(* IEC 61131-3 sources: daoli-st-library/DL_Device (part 17) *)

(* ---- FB_DL_CombinerArcDetect.st ---- *)
(*
  FB_DL_CombinerArcDetect  —  汇流箱直流拉弧特征判据 / Combiner box DC arc feature detection
  分类 Category : DL_Device
  码位 Code     : 16#03_2_00
  版本 Version  : 1.0.1
  溯源 Source   : NAMUR NE107 语义借鉴 · clean-room 实现，仅借分类/参数域/命名，未复制源码
  修订 Revision : v1.0.1 (R34 终审抽检) — ① 段 1 复位只清组态码 16#0002_0300，不再连带清 16#0002_0310
                  （原「无条件清锁存」使拉弧仍在时 bError 掉为 FALSE、uErrorId 归 0，而 eNe107 仍报 eFailure，
                  故障位/事件码/NE107 三者不同步，且 eAlarm 解除需第二次复位沿）；
                  ② bCfgOk 补 tSampleTime / tFilterTC 正域闸（原 0 或负值时高通静默不动作、永不告警，违 R179）。
                  接口、码表、NE107 映射不变。
  功能 Function : 1) 高通滤波提取电流高频分量，超门限按多拍持续确认才升故障（单拍尖峰只计信息级）；
                  2) 采样率与滤波截止频率配比校验（截止 >= 采样率/2 即出厂报码，不进入判据）；
                  3) 分级出口按 NE107 六态映射，未知态归 eUnknown 绝不归 eOk。
  边界 Boundary : ① 高频分量提取前确认采样率/截止频率配比合法（截止 >= 采样率/2 即报码）；
                  ② 拉弧判据多拍持续确认，单拍尖峰只计信息级不升故障；
                  ③ 分级出口按 NE107 六态映射，未知态归 eUnknown（不归 eOk）；
                  ④ 输出三行同向：高频分量 → 确认计数 → 拉弧标志。
  依赖 Depends  : FB_DL_HighPassFilter（高频分量提取，每拍无条件调用）

  码表 Error codes（本件子码步进 16#10，避让邻件码位）:
    16#0002_0300 故障级：采样率/截止频率配比非法（截止 >= 采样率/2）或采样率 <= 0
    16#0002_0310 故障级：拉弧已确认（多拍持续超门限），需 bReset 清除
    16#0002_0320 信息级：单拍尖峰（未达确认拍数，不置 bError）
*)

TYPE E_DL_CadNe107 :
(
    eOk                  := 0,   // 正常 / Normal
    eFailure             := 10,  // 故障 / Failure
    eCheckFunction       := 20,  // 功能检查 / Function check
    eOutOfSpec           := 30,  // 超出规格 / Out of specification
    eMaintenanceRequired := 40,  // 需要维护 / Maintenance required
    eUnknown             := 90   // 未知态（兜底）/ Unknown fallback
);
END_TYPE

TYPE E_DL_CadPhase :
(
    eIdle    := 0,   // 空闲 / Idle
    eWatch   := 10,  // 常规监视 / Normal watch
    eConfirm := 20,  // 多拍确认中 / Multi-scan confirmation
    eAlarm   := 30,  // 拉弧告警 / Arc alarm
    eFault   := 90   // 组态故障锁定 / Configuration fault locked
);
END_TYPE

FUNCTION_BLOCK FB_DL_CombinerArcDetect
VAR_INPUT
    bEnable       : BOOL;                         // 总使能，FALSE 回空闲 / Master enable
    bReset        : BOOL;                          // 复位，上升沿清告警与故障 / Reset
    fCurrentA     : REAL;                         // 直流支路电流 [A]，域 0~30 / DC branch current [A]
    fSampleRateHz : REAL := 10000.0;              // 电流采样率 [Hz]，域 > 0 / Current sampling rate [Hz]
    fCutoffHz     : REAL := 2000.0;               // 高通截止频率 [Hz]，须 < 采样率/2 / High-pass cutoff [Hz]
    fHfThreshA    : REAL := 0.15;                 // 高频分量门限 [A]，域 > 0 / HF component threshold [A]
    nConfirmScans : INT := 5;                     // 持续确认拍数 [拍]，域 1~100 / Confirmation scans, 1..100
    tFilterTC      : TIME := T#20MS;              // 高通时间常数 [ms] / High-pass time constant [ms]
    tSampleTime   : TIME := T#10MS;               // 任务采样周期 [ms]，域 > 0 / Task sample period [ms]
    fEps          : REAL := 1.0E-6;               // 浮点判零容差 [1] / Floating zero tolerance
END_VAR
VAR_OUTPUT
    fHfOutA       : REAL;                         // 高频分量输出 [A] / HF component output [A]
    nConfirmCnt   : INT;                          // 当前确认计数 [拍] / Current confirmation counter
    bArcAlarm     : BOOL;                         // 拉弧告警（保持型）/ Arc alarm, held
    bSpikeOnly    : BOOL;                         // 仅单拍尖峰（信息级）/ Single-scan spike only
    eNe107        : E_DL_CadNe107;                // NE107 六态映射出口，段尾单点赋值 / NE107 mapping, single write
    bError        : BOOL;                         // 故障标志，与故障级码配对 / Fault flag paired with fault codes
    uErrorId      : UDINT;                        // 事件码，0 = 无事件 / Event code, 0 = none
    eStateOut     : E_DL_CadPhase;                // 状态机当前态，段尾单点映射 / Phase mapped at tail
END_VAR
VAR
    _eState       : E_DL_CadPhase := E_DL_CadPhase.eIdle;  // 内部状态 / Internal state
    rtrReset      : R_TRIG;                       // 复位沿 / Reset edge
    fbHp          : FB_DL_HighPassFilter;         // 高通滤波实例（无条件调用）/ High-pass filter instance
    bCfgOk        : BOOL;                         // 配比组态合法 / Ratio configuration valid
    bSigOk        : BOOL;                         // 电流采样有效 / Current sample valid
    bOver         : BOOL;                         // 本拍超门限 / Over threshold this scan
    nCnt          : INT;                          // 确认计数暂存 [拍] / Confirmation counter buffer
    eMap          : E_DL_CadNe107;                // NE107 映射暂存（单点写入源）/ NE107 mapping buffer
    uFault        : UDINT;                        // 锁存故障码 / Latched fault code
    uInfo         : UDINT;                        // 信息级码 / Information code
END_VAR
VAR CONSTANT
    DL_CAD_CNTMAX : INT := 1000;                  // 确认计数上限 [拍]，防溢出 / Confirmation counter ceiling
    DL_CAD_SRMAX  : REAL := 1.0E6;                // 采样率物理域上限 [Hz] / Sampling rate domain high
END_VAR

(* === 段 0 · 实例刷新（无条件周期调用）=== *)
rtrReset(CLK := bReset);                          // 每拍刷新复位沿

(* === 段 1 · 组态闸：采样率/截止频率配比（截止 >= 采样率/2 即报码）=== *)
bCfgOk := (fSampleRateHz > fEps) AND (fSampleRateHz <= DL_CAD_SRMAX)
          AND (fCutoffHz > fEps)
          AND (fCutoffHz < (fSampleRateHz * 0.5))          // Nyquist 配比硬判据
          AND (fHfThreshA > fEps) AND (nConfirmScans >= 1) AND (nConfirmScans <= 100)
          AND (TIME_TO_LREAL(tSampleTime) > 0.0) AND (TIME_TO_LREAL(tFilterTC) > 0.0)   // 节拍/时间常数正域闸（R179）
          AND (fSampleRateHz = fSampleRateHz) AND (fCutoffHz = fCutoffHz)
          AND (fHfThreshA = fHfThreshA);                   // 含 NaN 自反判据
IF NOT bCfgOk THEN
    uFault := 16#0002_0300;                       // 故障级：配比非法
END_IF
IF rtrReset.Q AND bCfgOk THEN
    IF uFault <> 16#0002_0310 THEN
        uFault := 16#0000;                        // 复位沿清锁存（拉弧码由 eAlarm 相专清，保持位码同步）
    END_IF
    IF NOT bArcAlarm THEN
        nCnt := 0;                                // 未进入告警时清确认计数
    END_IF
END_IF
bSigOk := (fCurrentA = fCurrentA) AND (ABS(fCurrentA) < 1.0E30) AND (fCurrentA >= 0.0);   // NaN 自反 + 域闸
uInfo := 16#0000;                                 // 信息码每拍清零

(* === 段 2 · 高频分量实例（每拍无条件调用）=== *)
fbHp(bEnable := bEnable AND bSigOk AND bCfgOk,    // 配比非法/信号无效时不使能（禁误判）
     fIn := fCurrentA,                            // 电流采样
     tTimeConst := tFilterTC,                     // 高通时间常数
     tSampleTime := tSampleTime,                  // 采样周期
     rOutMin := -1000.0,                          // 输出下限 [A]
     rOutMax := 1000.0,                           // 输出上限 [A]
     bTrack := rtrReset.Q,                        // 复位沿清基线
     fTrackValue := 0.0);                         // 跟踪值 0
fHfOutA := fbHp.fOut;                             // 高频分量输出
bOver := bCfgOk AND bSigOk AND fbHp.bValid AND (ABS(fHfOutA) >= fHfThreshA);   // 超门限判据

(* === 段 3 · 主状态机（ENUM + CASE，含 ELSE 兜底）=== *)
CASE _eState OF
E_DL_CadPhase.eIdle :
    nCnt := 0;                                    // 空闲计数清零
    bSpikeOnly := FALSE;                          // 尖峰标志复位
    IF uFault = 16#0002_0300 THEN
        _eState := E_DL_CadPhase.eFault;          // 组态故障优先
    ELSIF bEnable AND bCfgOk THEN
        _eState := E_DL_CadPhase.eWatch;          // 进入监视相
    END_IF

E_DL_CadPhase.eWatch :
    IF bOver THEN
        nCnt := 1;                                // 首拍超门限：进入确认
        _eState := E_DL_CadPhase.eConfirm;
    ELSE
        IF bSpikeOnly THEN
            uInfo := 16#0002_0320;                // 信息级：单拍尖峰记录（不升故障）
        END_IF
        bSpikeOnly := bSpikeOnly AND bOver;       // 无超门限拍则尖峰记录清除
    END_IF

E_DL_CadPhase.eConfirm :
    IF bOver THEN
        nCnt := nCnt + 1;                         // 连续超门限：计数累加
        IF nCnt > DL_CAD_CNTMAX THEN
            nCnt := DL_CAD_CNTMAX;                // 饱和防溢出
        END_IF
        IF nCnt >= nConfirmScans THEN
            bArcAlarm := TRUE;                    // 置位型：拉弧确认告警（段尾不清零）
            uFault := 16#0002_0310;               // 故障级：拉弧已确认
            _eState := E_DL_CadPhase.eAlarm;      // 转告警相
        END_IF
    ELSE
        bSpikeOnly := TRUE;                       // 未达确认拍数即回落：只计单拍尖峰
        uInfo := 16#0002_0320;                    // 信息级：单拍尖峰
        nCnt := 0;                                // 计数清零（要求连续）
        _eState := E_DL_CadPhase.eWatch;          // 回监视相
    END_IF

E_DL_CadPhase.eAlarm :
    bArcAlarm := TRUE;                            // 告警保持
    IF NOT bOver AND rtrReset.Q THEN
        uFault := 16#0000;                        // 超门限消失且复位沿：清锁存
        bArcAlarm := FALSE;                       // 告警解除（可到达的解除路径）
        nCnt := 0;                                // 计数清零
        _eState := E_DL_CadPhase.eWatch;
    END_IF

E_DL_CadPhase.eFault :
    nCnt := 0;                                    // 故障态计数清零
    bArcAlarm := FALSE;                           // 故障态不告警（配置错误优先）
    IF uFault = 16#0000 THEN
        _eState := E_DL_CadPhase.eIdle;           // 解锁回空闲
    END_IF

ELSE
    _eState := E_DL_CadPhase.eFault;              // 非法状态拦截
    uFault := 16#0002_0300;                       // 故障级：相 ID 越界
    bArcAlarm := FALSE;                           // 安全侧不告警
END_CASE
IF NOT bEnable THEN
    _eState := E_DL_CadPhase.eIdle;               // 失能最高优先回空闲
    bArcAlarm := FALSE;                           // 失能清告警
    nCnt := 0;                                    // 失能清计数
    IF uFault = 16#0002_0310 THEN
        uFault := 16#0000;                        // 失能同拍清拉弧锁存：相序丢失后 eAlarm 不可达，防锁死（终审式 1）
    END_IF
END_IF

(* === 段 4 · 输出映射与 NE107 六态（段尾单点赋值）=== *)
nConfirmCnt := nCnt;                              // 确认计数输出
CASE _eState OF
E_DL_CadPhase.eWatch :
    eMap := E_DL_CadNe107.eOk;                    // 常规监视：正常态
E_DL_CadPhase.eConfirm :
    eMap := E_DL_CadNe107.eMaintenanceRequired;   // 确认中：需维护关注
E_DL_CadPhase.eAlarm :
    eMap := E_DL_CadNe107.eFailure;               // 拉弧确认：故障态
E_DL_CadPhase.eFault :
    eMap := E_DL_CadNe107.eOutOfSpec;             // 组态越规格
E_DL_CadPhase.eIdle :
    eMap := E_DL_CadNe107.eCheckFunction;         // 空闲未监视：功能检查
ELSE
    eMap := E_DL_CadNe107.eUnknown;               // 未知态兜底：绝不归 eOk
END_CASE
IF bSpikeOnly AND (eMap = E_DL_CadNe107.eOk) THEN
    eMap := E_DL_CadNe107.eMaintenanceRequired;   // 单拍尖峰：提升到需维护（信息级）
END_IF
eNe107 := eMap;                                   // 单点写入 NE107 出口
bError := (uFault <> 16#0000);                    // 故障标志仅由故障级码置位（R45 配对）
IF bError THEN
    uErrorId := uFault;                           // 故障级优先上报
ELSE
    uErrorId := uInfo;                            // 否则上报信息级码
END_IF
eStateOut := _eState;                             // 输出枚举段尾单点映射（N2 规则）
END_FUNCTION_BLOCK

(* ---- FB_DL_CondensateDrainSeq.st ---- *)
(*
  ==================================================================
  组件名 Component  : FB_DL_CondensateDrainSeq
  分类   Category   : DL_Device
  复杂度 Complexity  : cx5
  版本   Version    : 1.0.0
  功能   Purpose    : 储气罐 / 空压机冷凝水自动排污阀时序。定时触发与液位高
                      双触发源并联起排；开阀确认反馈 → 排放（触发消失且最
                      小排放时长满足）→ 关阀确认反馈；三窗超时诊断（开阀 /
                      排放 / 关阀独立成因独立码位语义，R190）。
  来源   Source     : t2-2-lbp（命令→监视→判定三段）
  溯源   Origin     : IEC 61131-3 标准语义的道莅防御性实现；冷凝水排污双触
                      发与阀反馈确认窗为行业公知工程语义，clean-room 自研实
                      现，未复制 LBP 或任何厂商私有库源码。
  平台   Platform   : 纯 IEC 61131-3（Standard.library: TON / R_TRIG，无私有库）
  分工声明 Split     : 与 DL_Device 存量阀类执行件（电磁阀直控类）分工——直
                      控件只做单阀开关映射，本件为排污全过程顺控（三窗监视
                      与诊断）；不做压力 / 温度工艺调节。
  作者   Author     : 道莅代码库 · PLC 编程专家（R58）
  ------------------------------------------------------------------
  边界 Boundary     :
                      一 组态配比约束（R100）：tMinDrain < tDrainMax（最小排
                         放短于排放超时）且 tOpenConfirm > T#0S 且 tCloseConfirm
                         > T#0S；越域判故障级锁存；
                      二 触发为电平语义：定时触发与液位高任一为真且许可满
                         足即起排；排放相退出 = 触发消失（事件）AND 最小排放
                         时长满足（双条件，R98 精神）；
                      三 故障相阀命令安全侧断开（排污阀断电 = 关闭，R191 显
                         式声明）；故障锁存解除路径 = bReset 上升沿（唯一路
                         径，R188）；
                      四 无全局变量、无外部变量声明、无物理地址寻址。
  修订记录 Revision  :
    2026-11-21  v1.0.0  R58 首版（批 3 · 序号 11）
  ==================================================================
*)

TYPE E_DL_CdsPhase :
(
    eCdsIdle    := 0,  // 空闲：等触发 / idle, waiting for a trigger
    eCdsOpening := 10, // 开阀：等阀开反馈确认 / opening, awaiting the open feedback
    eCdsDraining := 20, // 排放中：等触发消失且最小时长满足 / draining, awaiting the trigger gone with the minimum met
    eCdsClosing := 30, // 关阀：等阀关反馈确认 / closing, awaiting the closed feedback
    eCdsFault   := 90  // 故障锁存 / the latched fault
);
END_TYPE

TYPE E_DL_CdsCause :
(
    eNone         := 0, // 无成因 / no cause
    eCfgBad       := 1, // 组态非法：时间窗配比越域（故障级，与 bError 配对）/ an illegal config
    eValveOpenTo  := 2, // 开阀确认超时（故障级，与 bError 配对）/ an open confirm timeout
    eDrainTimeout := 3, // 排放超时（液位不回落，故障级，与 bError 配对）/ a drain timeout
    eValveCloseTo := 4, // 关阀确认超时（故障级，与 bError 配对）/ a close confirm timeout
    ePhaseBad     := 5  // 非法相位兜底（故障级，与 bError 配对）/ an illegal phase fallback
);
END_TYPE

FUNCTION_BLOCK FB_DL_CondensateDrainSeq
VAR_INPUT
    bEnable       : BOOL := TRUE;   // 使能，失能回空闲关阀 [-] / enable, disabling returns idle with the valve closed
    bReset        : BOOL := FALSE;  // 复位上升沿清故障锁存 [-] / reset rising edge clears the latch
    bTimTrig      : BOOL := FALSE;  // 定时触发电平（调用方定时器给出）[-] / the timer trigger level
    bLevelHigh    : BOOL := FALSE;  // 液位高触发电平 [-] / the level high trigger level
    bPermitDrain  : BOOL := TRUE;   // 排放许可（压力低联锁给出）[-] / the drain permit from the pressure interlock
    bFbValveOpen  : BOOL := FALSE;  // 排污阀开到位反馈 [-] / the valve open feedback
    bFbValveClosed: BOOL := TRUE;   // 排污阀关到位反馈 [-] / the valve closed feedback
    tOpenConfirm  : TIME := T#5S;   // 开阀确认窗 [毫秒] / the open confirm window [millisecond]
    tDrainMax     : TIME := T#60S;  // 排放超时窗 [毫秒] / the drain timeout window [millisecond]
    tCloseConfirm : TIME := T#5S;   // 关阀确认窗 [毫秒] / the close confirm window [millisecond]
    tMinDrain     : TIME := T#2S;   // 最小排放时长 [毫秒] / the minimum drain duration [millisecond]
END_VAR
VAR_OUTPUT
    bValveCmd   : BOOL := FALSE; // 排污阀命令输出（TRUE = 开阀）[-] / the valve command outlet, true = open
    bDrainActive: BOOL := FALSE; // 排放进行指示 [-] / the drain active indicator
    ePhase      : E_DL_CdsPhase := E_DL_CdsPhase.eCdsIdle; // 相位出口 [枚举] / the phase outlet
    eCause      : E_DL_CdsCause := E_DL_CdsCause.eNone; // 成因出口，锁存回放 [枚举] / the cause outlet replayed
    bError      : BOOL := FALSE; // 故障锁存标志 [-] / the fault latch flag
END_VAR
VAR
    rtReset : R_TRIG; // 复位沿检测，段 0 无条件刷新 / the reset edge
    tonOpen : TON;    // 开阀确认窗，段 0 无条件刷新 / the open confirm window
    tonDrain: TON;    // 排放超时窗，段 0 无条件刷新 / the drain timeout window
    tonClose: TON;    // 关阀确认窗，段 0 无条件刷新 / the close confirm window
    tonMin  : TON;    // 最小排放窗，段 0 无条件刷新 / the minimum drain window
    _ePhase : E_DL_CdsPhase := E_DL_CdsPhase.eCdsIdle; // 内部相位，CASE 唯一写入目标 / the internal phase
    _eFaulC : E_DL_CdsCause := E_DL_CdsCause.eNone; // 故障级成因，锁存至复位沿 / the fault cause latched
    _bFault : BOOL := FALSE; // 故障锁存位 [-] / the fault latch bit
    _bCfgOk : BOOL := FALSE; // 组态域内 [-] / the config inside the domain
    _bInit  : BOOL := FALSE; // 首扫初始化完成标志（R310）/ the first scan flag
END_VAR

// 段 0｜定时器与沿检测无条件周期刷新（禁入分支，FB50-1）/ segment 0, the unconditional refresh
rtReset(CLK := bReset); // 复位沿 / the reset edge
tonOpen(IN := (_ePhase = E_DL_CdsPhase.eCdsOpening) AND (NOT _bFault) AND bEnable, PT := tOpenConfirm); // 开阀窗，IN 串开阀相闸 / the open window gated by the opening phase
tonDrain(IN := (_ePhase = E_DL_CdsPhase.eCdsDraining) AND (NOT _bFault) AND bEnable, PT := tDrainMax); // 排放窗，IN 串排放相闸 / the drain window gated by the draining phase
tonClose(IN := (_ePhase = E_DL_CdsPhase.eCdsClosing) AND (NOT _bFault) AND bEnable, PT := tCloseConfirm); // 关阀窗，IN 串关阀相闸 / the close window gated by the closing phase
tonMin(IN := (_ePhase = E_DL_CdsPhase.eCdsDraining) AND (NOT _bFault) AND bEnable, PT := tMinDrain); // 最小排放窗，与排放窗同相起算（配比约束见边界一）/ the minimum window co-started with the drain window

// 段 1｜首扫初始化（R310）/ segment 1, the first scan
IF NOT _bInit THEN // 首扫一拍 / the first scan
    _bInit := TRUE; // 置首扫标志 / raise the flag
END_IF

// 段 2｜复位沿作用域：清故障锁存 / 迁空闲（两项逐项声明，边界三）/ segment 2, the reset edge scope
IF rtReset.Q THEN // 复位沿 / the reset edge
    _bFault := FALSE; // 作用域一：清故障锁存 / scope one, clear the fault latch
    _eFaulC := E_DL_CdsCause.eNone; // 作用域一：清成因 / scope one, clear the cause
    _ePhase := E_DL_CdsPhase.eCdsIdle; // 作用域二：迁空闲相 / scope two, back to idle
END_IF

// 段 3｜组态域闸（边界一，R100 配比）/ segment 3, the config gate
_bCfgOk := (tOpenConfirm > T#0S) AND (tCloseConfirm > T#0S) AND (tMinDrain < tDrainMax) AND (tDrainMax > T#0S); // 确认窗 / 排放窗 / 配比判定 / the confirm, drain and pairing verdicts
IF NOT _bCfgOk THEN // 配比越域 / a pairing violation
    IF NOT _bFault THEN // 未锁存才迁移 / migrate only while unlatched
        _bFault := TRUE; // 置故障锁存 / raise the fault latch
        _eFaulC := E_DL_CdsCause.eCfgBad; // 故障级成因（R45 配对）/ the fault cause
        _ePhase := E_DL_CdsPhase.eCdsFault; // 迁故障相（锁存与迁相同分支，FB50-1）/ migrate to the fault phase
    END_IF
END_IF

// 段 4｜相位机：ENUM + CASE，含 ELSE 非法相位兜底（R128）/ segment 4, the phase machine
CASE _ePhase OF

E_DL_CdsPhase.eCdsIdle: // 空闲相：双触发源并联评估（边界二）/ the idle phase, the dual trigger evaluation
    IF NOT bEnable THEN // 失能驻留 / dwell while disabled
        _ePhase := E_DL_CdsPhase.eCdsIdle; // 停摆驻留 / dwell
    ELSIF (bTimTrig OR bLevelHigh) AND bPermitDrain THEN // 触发且许可 / a trigger with the permit
        _ePhase := E_DL_CdsPhase.eCdsOpening; // 迁开阀相 / migrate to the opening phase
    END_IF

E_DL_CdsPhase.eCdsOpening: // 开阀相：等阀开反馈确认 / the opening phase
    IF NOT bEnable THEN // 失能回空闲关阀（R191 显式）/ a disable returns idle
        _ePhase := E_DL_CdsPhase.eCdsIdle; // 回空闲相 / back to idle
    ELSIF bFbValveOpen THEN // 阀开反馈确认 / the open feedback confirmed
        _ePhase := E_DL_CdsPhase.eCdsDraining; // 迁排放相 / migrate to the draining phase
    ELSIF tonOpen.Q THEN // 开阀确认窗超时（R190 独立成因）/ the open timeout, an independent cause
        _bFault := TRUE; // 置故障锁存 / raise the fault latch
        _eFaulC := E_DL_CdsCause.eValveOpenTo; // 故障级成因（R45 配对）/ the fault cause
        _ePhase := E_DL_CdsPhase.eCdsFault; // 迁故障相 / migrate to the fault phase
    END_IF

E_DL_CdsPhase.eCdsDraining: // 排放相：双退出条件（边界二，R98 精神）/ the draining phase, the dual exit
    IF NOT bEnable THEN // 失能回空闲关阀 / a disable returns idle
        _ePhase := E_DL_CdsPhase.eCdsIdle; // 回空闲相 / back to idle
    ELSIF (NOT bTimTrig) AND (NOT bLevelHigh) AND tonMin.Q THEN // 触发消失且最小排放时长满足 / the trigger gone with the minimum met
        _ePhase := E_DL_CdsPhase.eCdsClosing; // 迁关阀相 / migrate to the closing phase
    ELSIF tonDrain.Q THEN // 排放超时（液位不回落，R190 独立成因）/ the drain timeout, an independent cause
        _bFault := TRUE; // 置故障锁存 / raise the fault latch
        _eFaulC := E_DL_CdsCause.eDrainTimeout; // 故障级成因（R45 配对）/ the fault cause
        _ePhase := E_DL_CdsPhase.eCdsFault; // 迁故障相 / migrate to the fault phase
    END_IF

E_DL_CdsPhase.eCdsClosing: // 关阀相：等阀关反馈确认 / the closing phase
    IF NOT bEnable THEN // 失能回空闲 / a disable returns idle
        _ePhase := E_DL_CdsPhase.eCdsIdle; // 回空闲相 / back to idle
    ELSIF bFbValveClosed THEN // 阀关反馈确认 / the closed feedback confirmed
        _ePhase := E_DL_CdsPhase.eCdsIdle; // 回空闲相 / back to idle
    ELSIF tonClose.Q THEN // 关阀确认窗超时（R190 独立成因）/ the close timeout, an independent cause
        _bFault := TRUE; // 置故障锁存 / raise the fault latch
        _eFaulC := E_DL_CdsCause.eValveCloseTo; // 故障级成因（R45 配对）/ the fault cause
        _ePhase := E_DL_CdsPhase.eCdsFault; // 迁故障相 / migrate to the fault phase
    END_IF

E_DL_CdsPhase.eCdsFault: // 故障相：成因锁存等复位沿；阀命令安全侧断开 / the fault phase
ELSE // 非法相位兜底（R128）/ the illegal phase fallback
    _bFault := TRUE; // 置故障锁存 / raise the fault latch
    _eFaulC := E_DL_CdsCause.ePhaseBad; // 故障级成因（R45 配对）/ the fault cause
    _ePhase := E_DL_CdsPhase.eCdsFault; // 迁故障相 / migrate to the fault phase
END_CASE

// 段 5｜统一出口（边界三安全侧）/ segment 5, the unified outlet
bValveCmd := ((_ePhase = E_DL_CdsPhase.eCdsOpening) OR (_ePhase = E_DL_CdsPhase.eCdsDraining)) AND bEnable AND (NOT _bFault); // 阀命令仅开阀与排放相 / the valve command in the opening and draining phases
bDrainActive := (_ePhase = E_DL_CdsPhase.eCdsDraining) AND (NOT _bFault); // 排放指示 / the drain indicator
ePhase := _ePhase; // 相位出口单点映射 / the phase outlet
IF _bFault THEN // 故障锁存优先 / the fault latch first
    eCause := _eFaulC; // 成因锁存回放（R152）/ the cause replayed
ELSE // 无锁存 / no latch
    eCause := E_DL_CdsCause.eNone; // 无成因 / no cause
END_IF
bError := _bFault; // 故障标志与锁存位同源 / the flag shares the latch
END_FUNCTION_BLOCK

(* ---- FB_DL_ContactorWeldDetect.st ---- *)
(*==============================================================================
 * 组件名称 (Component)  : FB_DL_ContactorWeldDetect
 * 所属子库 (Sublibrary) : DL_Device
 * 当前版本 (Version)    : 1.0.0
 * 兼容性   (Platform)   : CODESYS 3.5+ / TwinCAT 3 / 汇川 InoProShop / 施耐德 Machine Expert
 *                         仅依赖 Standard.library（TON / R_TRIG）与库内健康枚举唯一属主，
 *                         零厂商私有库
 * 功能描述 (Function)   : 接触器熔焊与不吸合检测。① 熔焊：断开指令后 tReleaseMax 内反馈仍为 1
 *                         → eCause = eWeld，故障锁存；② 不吸合：闭合指令后 tPickupMax 内无反馈
 *                         → eCause = eNoPickup，故障锁存。两成因各有独立 TON 与独立归因成员
 *                         （R190 归因唯一，禁止共用一个成因导致另一端永不赋值）。
 * 复位语义 (Design)     : **熔焊为不可自恢复故障**：解除式要求「复位沿 ∧ 反馈已回落」。若反馈是
 *                         真实熔焊，反馈不会回落 → 复位**不解锁**，这是**设计意图**而非缺陷：
 *                         触点焊死时允许软复位等于给现场一个「假修复」通道，会把带电粘连的
 *                         主回路重新投入。现场处置只能是更换接触器后反馈自然回落再复位。
 * 归属声明 (Ownership)  : 健康出口 eHealth 引用枚举 `E_DL_Ne107Status` 唯一属主，属主文件为
 *                         `C:\Library\DL_Device\I_DL_DeviceHealth.st`（枚举定义位于该文件 L91 附近），
 *                         本件只引用不重复声明（全库同名枚举定义计数 = 1，R67）。
 * 接口     (Interface)  : 输入 bCmdClose 闭合指令、bFbClosed 触点反馈、tReleaseMax 释放超时、
 *                         tPickupMax 吸合超时、bReset 复位；输出 bWeldSuspect 熔焊疑似位、
 *                         eCause 归因、eHealth NE107 健康态、eState / bError / nErrId。
 * 边界     (Boundary)   : ① 组态闸：tReleaseMax <= T#0S 或 tPickupMax <= T#0S → 故障锁存；
 *                         ② TON 两枚 + R_TRIG 一枚段 0 无条件周期刷新，IN 由当拍指令与反馈派生；
 *                         ③ 故障相迁出唯一路径 = bReset 上升沿；④ 零全局耦合（无 GVL / 无物理地址）。
 * 解除式   (Release)    : bReset 上升沿 ∧ 组态合法 ∧ 反馈已回落（bFbClosed = FALSE，当拍量，
 *                         R240 范式）。自证可满足（终审两式 1）：反馈为真实熔焊时该式不可满足，
 *                         属刻意的安全不可解除；触点更换后反馈回落即达，故路径物理可达。
 * 码表     (Codes)      : 16#0003_0702 故障级：接触器故障总码（组态非法 / 熔焊 / 不吸合 / 非法相位），
 *                         锁存至 bReset 上升沿，归因由 eCause 承载（R190 单件单总码）；
 *                         16#0003_0481 信息级：吸合动作正常确认（指令闭合且反馈已到位）。
 *                         加码反证（R90）：吸合正常确认与「一直闭合保持着」在 bFbClosed / bError 上
 *                         完全同值，出口组合无法区分「刚完成一次吸合确认」与「长期闭合」，
 *                         故立一码留痕。
 *                         码段说明：Device 的 03xx 故障子带已占满（仅余 03C5~03C9 碎片孔洞，按
 *                         实战规则 13 禁回填），故本批新开 07xx 故障子带取 16#0003_0702；
 *                         信息级用 04xx 子带取 16#0003_0481（源码实扫为空）。分段理由即此。
 * 开源溯源 (Origin)     : 道莅自研 clean-room（参考设备级 AOI 熔焊检测粒度与参数域，
 *                         零代码行复制；t2-6-rockwell-aoi 族）
 * 修订历史 (Revision)   : 2026-11-19  v1.0.0  R45 首版（批次 4 · 序号 16）
 *==============================================================================*)

TYPE E_DL_CwdState :
(
    eIdle  := 0,     // 待机（指令与反馈均断开） / Idle, command and feedback both released
    eRun   := 10,    // 动作监视 / Monitoring motion
    eFault := 90     // 故障锁存相 / Fault latched phase
);
END_TYPE

TYPE E_DL_CwdCause :
(
    eNone       := 0,   // 无故障成因 / No cause
    eCfgIllegal := 1,   // 组态非法 / Illegal configuration
    eWeld       := 2,   // 熔焊（断开指令后反馈不回落） / Welded, feedback stays on after release
    eNoPickup   := 3,   // 不吸合（闭合指令后无反馈） / No pickup, no feedback after close
    ePhaseBad   := 4    // 非法相位兜底 / Illegal phase fallback
);
END_TYPE

FUNCTION_BLOCK FB_DL_ContactorWeldDetect
VAR_INPUT
    bCmdClose    : BOOL := FALSE;        // 闭合指令 [-] / Close command
    bFbClosed    : BOOL := FALSE;        // 主/辅助触点反馈（TRUE = 已闭合） [-] / Contact feedback, TRUE means closed
    tReleaseMax  : TIME := T#500MS;      // 释放允许时间，域 > T#0S [ms] / Release allowance, domain > T#0S [ms]
    tPickupMax   : TIME := T#300MS;      // 吸合允许时间，域 > T#0S [ms] / Pickup allowance, domain > T#0S [ms]
    bReset       : BOOL := FALSE;        // 复位命令，上升沿清故障（真实熔焊时不解锁为设计意图） [-] / Reset, does not unlock a truly welded contact by design
END_VAR
VAR_OUTPUT
    bWeldSuspect : BOOL;                 // 熔焊疑似（锁存回放） [-] / Weld suspect, latched replay
    eCause       : E_DL_CwdCause;        // 故障成因出口（R190 归因唯一） / Fault cause outlet
    eHealth      : E_DL_Ne107Status;     // NE107 健康态（引用唯一属主枚举） [-] / NE107 health, owner enum referenced
    eState       : E_DL_CwdState;        // 状态出口，段 6 单点映射 / State outlet
    bError       : BOOL;                 // 故障锁存标志 [-] / Fault latch flag
    nErrId       : UDINT;                // 事件码，0 = 无事件 / Event code, 0 = no event
END_VAR
VAR
    _eState      : E_DL_CwdState := E_DL_CwdState.eIdle;     // 内部相位（CASE 唯一写入目标） / Internal phase
    _eCause      : E_DL_CwdCause := E_DL_CwdCause.eNone;     // 故障成因锁存（锁存量） / Latched cause
    tonRelease   : TON;                  // 释放超时计时，段 0 无条件调用 / Release timeout timer
    tonPickup    : TON;                  // 吸合超时计时，段 0 无条件调用 / Pickup timeout timer
    rtReset      : R_TRIG;               // 复位沿实例，段 0 无条件调用 / Reset edge
    _bWeldLatch  : BOOL;                 // 熔焊疑似锁存位（锁存量） / Weld suspect latch
    _bCfgBad     : BOOL;                 // 组态非法当拍量 [-] / Illegal configuration
    _bFault      : BOOL;                 // 故障锁存位（锁存量） / Latched fault bit
    _uFault      : UDINT;                // 故障码锁存（锁存量） / Latched fault code
    _uInfo       : UDINT;                // 信息码，每拍重算 / Info code, recomputed each scan
END_VAR

(* —— 段 0：当拍判据派生 + 定时器与沿实例无条件周期刷新 —— *)
_bCfgBad := (tReleaseMax <= T#0S) OR (tPickupMax <= T#0S);                                // 组态域闸 / Configuration gate
rtReset(CLK := bReset);                                                                   // 复位沿，每拍必调（R228A） / Reset edge
tonRelease(IN := (NOT bCmdClose) AND bFbClosed, PT := tReleaseMax);                        // 释放超时计时（断开后反馈仍在） / Release timeout
tonPickup(IN := bCmdClose AND (NOT bFbClosed), PT := tPickupMax);                          // 吸合超时计时（闭合后无反馈） / Pickup timeout

(* —— 段 1：单拍量预清零（锁存量不入清单，R107） —— *)
_uInfo       := 16#0000_0000;      // 信息码每拍重算 / Info recomputed every scan
bWeldSuspect := FALSE;             // 熔焊疑似位缺省假，由锁存回放 / Weld suspect preset
nErrId       := 16#0000_0000;      // 事件码缺省无事件 / Event code default none
bError       := FALSE;             // 故障标志每拍预清，故障分支同拍置位（R45 配对） / Flag preset

(* —— 段 2：复位沿 + 组态域闸 —— *)
IF rtReset.Q THEN                                                        // 当拍复位沿 / current-scan reset edge
    _bFault := FALSE;                                                    // 清故障锁存位（锁存量） / Clear fault latch
    _uFault := 16#0000_0000;                                             // 清故障锁存码（锁存量） / Clear latched code
    _eCause := E_DL_CwdCause.eNone;                                      // 清成因（锁存量） / Clear latched cause
    IF _eState = E_DL_CwdState.eFault THEN
        _eState := E_DL_CwdState.eIdle;                                  // 故障相迁出唯一路径 / Sole exit from fault phase
    END_IF
END_IF
IF _bCfgBad THEN                                                         // 组态域闸 / Configuration gate
    _uFault := 16#0003_0702;                                             // 故障级：接触器故障总码 / Fault-level: contactor fault code
    _bFault := TRUE;
    bError  := TRUE;                                                     // 故障标志同拍置位（R45 配对） / Error flag set same scan
    _eCause := E_DL_CwdCause.eCfgIllegal;                                // 归因：组态非法 / Cause: illegal configuration
END_IF

(* —— 段 3：熔焊 / 不吸合双判据（各用独立实例与独立归因，R190） —— *)
IF (NOT _bFault) AND tonRelease.Q THEN                                   // 熔焊判据：断开后反馈不回落 / Weld criterion
    _uFault := 16#0003_0702;
    _bFault := TRUE;
    bError  := TRUE;
    _eCause := E_DL_CwdCause.eWeld;                                      // 归因：熔焊 / Cause: welded
    _bWeldLatch := TRUE;                                                 // 熔焊疑似锁存（供 HMI 持续显示） / Latch weld suspicion
END_IF
IF (NOT _bFault) AND tonPickup.Q THEN                                    // 不吸合判据：闭合后无反馈 / No-pickup criterion
    _uFault := 16#0003_0702;
    _bFault := TRUE;
    bError  := TRUE;
    _eCause := E_DL_CwdCause.eNoPickup;                                  // 归因：不吸合 / Cause: no pickup
END_IF
IF (NOT _bFault) AND bCmdClose AND bFbClosed THEN                        // 吸合正常确认（信息级） / Normal pickup confirmed
    _uInfo := 16#0003_0481;
END_IF

(* —— 段 4：故障解除式（R240 全当拍量；真实熔焊不解锁为设计意图） —— *)
IF rtReset.Q AND (NOT _bCfgBad) AND (NOT bFbClosed) THEN
    _bFault := FALSE;                                                    // 清故障锁存位（锁存量） / Clear fault latch
    _uFault := 16#0000_0000;                                             // 清故障锁存码（锁存量） / Clear latched code
    _eCause := E_DL_CwdCause.eNone;                                      // 清成因（锁存量） / Clear latched cause
    _bWeldLatch := FALSE;                                                // 反馈已回落才撤熔焊疑似 / Clear weld suspicion only after feedback dropped
END_IF

(* —— 段 4A：故障锁存相位迁移闸 —— *)
IF _bFault AND (_eState <> E_DL_CwdState.eFault) THEN
    _eState := E_DL_CwdState.eFault;                                     // 锁存即入故障相 / Latch enters fault phase
END_IF

(* —— 段 5：相位机（ENUM 全成员显式标签 + ELSE 兜底，R128） —— *)
CASE _eState OF

E_DL_CwdState.eIdle:
    IF (bCmdClose OR bFbClosed) AND (NOT _bFault) THEN                   // 出口 1：出现动作 / Motion appears
        _eState := E_DL_CwdState.eRun;
    ELSIF _bFault THEN                                                   // 出口 2：故障锁存 / Fault latched
        _eState := E_DL_CwdState.eFault;
    END_IF

E_DL_CwdState.eRun:
    IF (NOT bCmdClose) AND (NOT bFbClosed) AND (NOT _bFault) THEN        // 出口 1：指令与反馈均已复原（前置消失，R98） / Both released
        _eState := E_DL_CwdState.eIdle;
    ELSIF _bFault THEN                                                   // 出口 2：故障锁存 / Fault latched
        _eState := E_DL_CwdState.eFault;
    END_IF

E_DL_CwdState.eFault:
    ;                                                                     // 故障相：仅段 4 复位沿可迁出 / Only the reset edge leaves this phase

ELSE
    _uFault := 16#0003_0702;                                             // 故障级：非法相位兜底（归并总码） / Illegal-phase fallback
    _bFault := TRUE;
    bError  := TRUE;
    _eCause := E_DL_CwdCause.ePhaseBad;                                  // 归因：非法相位 / Cause: illegal phase
    _eState := E_DL_CwdState.eFault;

END_CASE

(* —— 段 6：出口单点映射（名实同源；锁存码回放；NE107 健康态仲裁） —— *)
bWeldSuspect := _bWeldLatch AND _bFault;                                 // 熔焊疑似仅在故障锁存期成立（名实同源） / Weld suspicion only while latched
IF _bFault OR _bCfgBad THEN
    eHealth := E_DL_Ne107Status.eFailure;                                // 失效级 / Failure level
ELSIF bCmdClose AND (NOT bFbClosed) THEN
    eHealth := E_DL_Ne107Status.eCheckFunction;                          // 吸合动作确认中（信号暂不可信） / Function check during pickup
ELSE
    eHealth := E_DL_Ne107Status.eOk;                                     // 正常级 / OK level
END_IF
IF _bFault THEN
    nErrId := _uFault;                                                   // 故障锁存码回放 / Replay latched fault code
ELSE
    nErrId := _uInfo;                                                    // 信息码 / Info code
END_IF
bError := _bFault;                                                       // 故障标志与锁存同源（名实双出口，R191） / Flag from latch
eState := _eState;                                                       // 状态出口 / State outlet
eCause := _eCause;                                                       // 成因出口 / Cause outlet

END_FUNCTION_BLOCK

(* ---- FB_DL_ControlValveDiag.st ---- *)
(*==============================================================================
 * 组件名称 (Component)  : FB_DL_ControlValveDiag
 * 溯源说明 (Provenance) : 道莅 clean-room 防御性实现（LBP 深化，补调节阀诊断缺口）
 * 所属子库 (Sublibrary) : DL_Device / ValveDiag
 * 当前版本 (Version)    : 1.0.0
 * 兼容性   (Platform)   : CODESYS 3.5 / TwinCAT 3 / 汇川 InoProShop；
 *                         纯 IEC 61131-3（第 3 版），仅用标准库 TON / R_TRIG
 * 组件分类 (Category)   : 功能块（FUNCTION_BLOCK）· 调节阀行程偏差与迟滞诊断
 * 功能一句话 (Summary)  : 行程偏差确认 + 迟滞估计 + NE107 健康分级，仅监视不驱动。
 * 边界与安全 (Boundary) : ①反馈小于 -5% 或大于 105% → 传感器故障态优先于偏差态；
 *                         ②bEnable=FALSE → 全部输出复位（安全侧缺省）；
 *                         ③累计行程按反馈逐拍绝对增量累积（寿命估计口径）；
 *                         ④迟滞按指令换向点反馈快照对估计，超带锁存置码；
 *                         ⑤偏差 TON 与换向沿检测各一次、无条件周期刷新；
 *                         ⑥健康分级映射：传感器故障=eFailure，
 *                           偏差确认=eMaintenanceReq，迟滞超带=eOutOfSpec，
 *                           其余=eOk（数值小者即最严级，与库公约一致）。
 * 错误码    : 16#0003_0375 反馈超量程（传感器故障态）——故障级（持续态）
 *             16#0003_0376 行程偏差确认超时——故障级（持续态）
 *             16#0003_0377 迟滞超带（估计值大于容带）——故障级（持续态）
 * 码位总账  : 16#0003_0375 用 / 16#0003_0376 用 / 16#0003_0377 用
 * 修改记录  : v1.0.0 R26 初版
 *==============================================================================*)
FUNCTION_BLOCK FB_DL_ControlValveDiag
VAR_INPUT
    fCmdPos   : LREAL; // 指令阀位 [%] / Commanded valve position [%]
    fFbPos    : LREAL; // 反馈阀位 [%] / Feedback valve position [%]
    fDevLimit : LREAL; // 偏差容限 [%] / Deviation limit [%]
    tDevDelay : TIME;  // 偏差确认延时 [ms] / Deviation confirm delay [ms]
    fHystBand : LREAL; // 迟滞容带 [%] / Hysteresis band [%]
    bEnable   : BOOL;  // 监视使能 / Monitoring enable
END_VAR
VAR_OUTPUT
    eHealth        : E_DL_Ne107Status; // NE107 健康分级 / NE107 health classification
    bDeviationAlarm: BOOL; // 偏差确认告警 / Confirmed deviation alarm
    fDeviation     : LREAL; // 当前行程偏差 [%] / Current stroke deviation [%]
    uTravelAccum   : LREAL; // 累计行程 [%]（原规格非标类型按红线 2 改 LREAL）/ Accumulated travel [%]
    eErr           : UDINT; // 本周期错误码，0=无错 / Error code this cycle, 0 = none
END_VAR
VAR
    fFbPrev   : LREAL;  // 上拍反馈锁存（行程增量与方向判据源）/ Previous feedback latch
    bFbPrevOk : BOOL;   // 上拍反馈有效性（首拍防假增量）/ Previous feedback validity
    fDevAbs   : LREAL;  // 偏差绝对值 / Absolute deviation
    fDelta    : LREAL;  // 反馈逐拍增量临时量 / Feedback per-cycle delta temp
    tonDev    : TON;    // 偏差确认定时器（单实例无条件刷新）/ Deviation confirm timer
    rDirUp    : R_TRIG; // 指令下转上换向沿（单实例无条件刷新）/ Up-reversal edge
    rDirDn    : R_TRIG; // 指令上转下换向沿（单实例无条件刷新）/ Down-reversal edge
    iCmdDir   : INT;    // 本拍指令方向（1 上 / -1 下 / 0 平）/ Command direction this cycle
    iDirPrev  : INT;    // 上拍指令方向 / Previous command direction
    fSnapUp   : LREAL;  // 上行换向反馈快照 / Feedback snapshot at up-reversal
    bSnapUpOk : BOOL;   // 上行快照有效 / Up snapshot valid
    fHystEst  : LREAL;  // 迟滞估计值 [%] / Hysteresis estimate [%]
    bHystTripped: BOOL; // 迟滞超带锁存 / Hysteresis over-band latch
    fFbGuard  : LREAL;  // 反馈实时守卫副本（内部判定统一用）/ Live feedback guard copy
END_VAR

// ---------- 实时反馈守卫副本：内部判定统一用此副本（对外无副本输出） ----------
fFbGuard := fFbPos;

// ---------- 使能为假：全输出复位（安全侧缺省） ----------
IF NOT bEnable THEN
    eHealth         := E_DL_Ne107Status.eUnknown; // 未监视态 / Unknown when disabled
    bDeviationAlarm := FALSE;
    fDeviation      := 0.0;
    uTravelAccum    := 0.0;
    eErr            := 0;
    bFbPrevOk   := FALSE;                     // 重置首拍防假增量 / Reset first-scan guard
    bSnapUpOk   := FALSE;
    fHystEst    := 0.0;
    bHystTripped := FALSE;
    iDirPrev    := 0;
    // 定时器与沿检测仍在下方无条件刷新（IN 条件含使能，禁能即静止）/ Timers refreshed unconditionally below
ELSE
    // ---------- 行程偏差绝对值（先算后喂定时器，禁先行使用） ----------
    fDeviation := fCmdPos - fFbGuard;         // 实时偏差 / Live deviation
    fDevAbs    := fDeviation;
    IF fDevAbs < 0.0 THEN
        fDevAbs := -fDevAbs;                  // 手工取反绝对值 / Manual absolute value
    END_IF
END_IF

// ---------- 无条件周期刷新：偏差 TON 与双向换向沿（各仅一次） ----------
tonDev(IN := bEnable AND (fDevAbs > fDevLimit) AND (fFbGuard >= -5.0) AND (fFbGuard <= 105.0),
       PT := tDevDelay);

// ---------- 指令方向判定（相邻拍指令差） ----------
iCmdDir := 0;
IF fCmdPos > fFbPrev THEN
    iCmdDir := 1;                             // 上行 / Rising
ELSIF fCmdPos < fFbPrev THEN
    iCmdDir := -1;                            // 下行 / Falling
END_IF
rDirUp(CLK := (iCmdDir = 1) AND (iDirPrev = -1)); // 下转上换向 / Reversal down-to-up
rDirDn(CLK := (iCmdDir = -1) AND (iDirPrev = 1)); // 上转下换向 / Reversal up-to-down

// ---------- 使能门控的主判定（禁能时跳过诊断结论更新） ----------
IF bEnable THEN
    // ---------- 反馈超量程：传感器故障态优先于偏差态 ----------
    IF (fFbGuard < -5.0) OR (fFbGuard > 105.0) THEN
        eHealth := E_DL_Ne107Status.eFailure; // 传感器故障最严级 / Sensor fault strictest
        eErr    := 16#0003_0375;              // 超量程码 / Out-of-range code
        bDeviationAlarm := FALSE;             // 偏差态被覆盖 / Deviation overridden
        fDeviation := 0.0;
        bFbPrevOk := FALSE;                   // 量程外不累积行程 / No travel accumulation
    ELSE
        // ---------- 偏差确认 ----------
        IF tonDev.Q THEN
            bDeviationAlarm := TRUE;          // 偏差确认成立 / Deviation confirmed
            eErr := 16#0003_0376;             // 确认超时码 / Confirm code
        ELSE
            bDeviationAlarm := FALSE;         // 未确认即撤销 / Withdrawn if unconfirmed
        END_IF

        // ---------- 累计行程：反馈逐拍绝对增量（寿命估计口径） ----------
        IF bFbPrevOk THEN
            fDelta := fFbGuard - fFbPrev;     // 逐拍增量 / Per-cycle delta
            IF fDelta < 0.0 THEN
                fDelta := -fDelta;            // 绝对增量 / Absolute delta
            END_IF
            uTravelAccum := uTravelAccum + fDelta; // 累积行程 / Accumulate
        END_IF
        bFbPrevOk := TRUE;
        fFbPrev   := fFbGuard;                // 锁存本拍反馈 / Latch feedback

        // ---------- 迟滞估计：下行换向时与上行快照配对 ----------
        IF rDirUp.Q THEN
            fSnapUp   := fFbGuard;            // 上行换向快照 / Up-reversal snapshot
            bSnapUpOk := TRUE;
        END_IF
        IF rDirDn.Q AND bSnapUpOk THEN
            fHystEst := fSnapUp - fFbGuard;   // 快照对差值 / Snapshot pair difference
            IF fHystEst < 0.0 THEN
                fHystEst := -fHystEst;        // 绝对迟滞 / Absolute hysteresis
            END_IF
            IF fHystEst > fHystBand THEN
                bHystTripped := TRUE;         // 超带锁存（需禁能复位）/ Over-band latch
            END_IF
        END_IF

        // ---------- NE107 分级仲裁（数值小者最严） ----------
        IF bHystTripped THEN
            eHealth := E_DL_Ne107Status.eOutOfSpec;       // 迟滞超带 / Out of spec
            IF eErr = 0 THEN
                eErr := 16#0003_0377;         // 迟滞超带码（不覆盖更严码）/ Hysteresis code
            END_IF
        ELSIF bDeviationAlarm THEN
            eHealth := E_DL_Ne107Status.eMaintenanceReq;  // 偏差确认 / Maintenance required
        ELSE
            eHealth := E_DL_Ne107Status.eOk;  // 监视中无异常 / Monitored, healthy
        END_IF
    END_IF
END_IF

END_FUNCTION_BLOCK

(* ---- FB_DL_ConveyorJamDetect.st ---- *)
(*
    FB_DL_ConveyorJamDetect —— 输送线堵料检测（无件时长 + 电机电流 双判据）
    ------------------------------------------------------------------
    组件名称  : FB_DL_ConveyorJamDetect
    分类      : DL_Device / ConveyorDiagnostics
    前缀      : FB_DL_
    版本      : 1.0.0
    溯源      : 借鉴点 —— 输送线堵料的两条经典判据及其组合方式：其一下游长时间
                无件到达（物料流中断）、其二驱动电机电流偏高（负载增大），
                二者同时成立才判堵料（单一判据都会误报：无件也可能是上游空料，
                电流高也可能是启动冲击或低温黏滞）；电流侧带回差释放线，
                两侧均带独立延时确认。该组合判据为公开工程常识。
                clean-room 声明 —— 零代码行复制；判据结构、闸门、锁存、码位与
                双语文档全部本件自有，仅使用 IEC 61131-3 标准库 TON / R_TRIG。
                许可证 —— 本件 MIT；来源标签 self-std（道莅自有内规族）。
    平台      : 纯 IEC 61131-3，CODESYS 3.5 / TwinCAT 3 / InoProShop / Machine Expert 通用
    作者      : 道莅代码库 · PLC编程专家（R70 构建轮 · 批 2 · N7）
    ------------------------------------------------------------------
    功能说明  : 判据一（无件）：输送机在运行（bConvRun）且下游件检测（bDownPart）
                持续为 FALSE 达 tNoPart → 无件确认位 _tonNoPart.Q。
                判据二（电流）：fMotorA 超过 fCurrHigh 且持续 tConfirm → 电流确认位；
                释放线为 fCurrHigh - fCurrHyst（回差，取确认位的自保持在条件内实现，
                与 FB_DL_ScaleRangeWatch 采用同一口径，全库口径一致）。
                合成：两侧确认位同时成立 → 堵料锁存 _bJam，bReset 上升沿解除；
                解除后若两侧条件仍成立，需重新满足两个延时才会再次判堵
                （避免复位后立刻重锁）。
                判据优先级：堵料锁存 > 组态/输入故障码；故障期内不重推断成因（R189）。
    错误码    : 16#0002_0601 组态非法（阈值 / 回差 / 时长 / 非有限），锁存 —— 故障级
                16#0002_0602 电机电流非有限，锁存 —— 故障级
                16#0002_0603 堵料判定（双判据同时确认），锁存至 bReset —— 故障级
    码位总账  : 0601 / 0602 / 0603 用（均故障级）；无信息级码（bBusy / 各确认位已可观测）
    状态机    : N/A —— 无顺序相（两侧确认由 TON 自持，属定时器状态），
                故无 ENUM / CASE，也无 CASE ELSE 兜底面
    边界与披露: 一 组态闸（R272 逐项点名）：fCurrHigh > 0；fCurrHyst >= 0；
                   fCurrHyst < fCurrHigh（否则释放线为负，判据恒自保持）；
                   fCurrHigh / fCurrHyst 非有限闸（NaN 自反 + Inf 差值自反 + 幅值上界）；
                二 输入闸：fMotorA 非有限 → 锁存 0602，两侧确认位清零（不判堵）；
                三 出口语义（R191 名实双出口）：bJam 为**保持量**（锁存后保持 TRUE 直到
                   复位），bError 为 bJam 与故障锁存的并；失能（bEn = FALSE）时
                   bJam 保持量**不被清除**（失能非复位），但 bBusy 与各确认位清零；
                四 定时器 _tonNoPart / _tonConfirm 每周期无条件调用（规则 ⑦），
                   IN 为显式条件表达式，未放入任何可被跳过的分支；
                五 浮点判据全部为不等式（>、<、>=），无浮点直比；无除法；无数组下标；
                六 零全局变量、零 VAR_EXTERNAL、零物理地址。
    修订记录  : 2026-11-22 v1.0.0 首次入库（R70 构建轮 · 批 2 · N7）
*)
FUNCTION_BLOCK FB_DL_ConveyorJamDetect
VAR_INPUT
    bEn        : BOOL := TRUE;             (* 使能，[标志] / the enable *)
    bReset     : BOOL := FALSE;            (* 堵料复位（上升沿有效），[标志] / the jam reset, rising edge *)
    bConvRun   : BOOL := FALSE;            (* 输送机运行反馈，[标志] / the conveyor running feedback *)
    bDownPart  : BOOL := FALSE;            (* 下游件检测（有件为真），[标志] / the downstream part present *)
    fMotorA    : LREAL := 0.0;             (* 驱动电机电流，[A] / the drive motor current *)
    fCurrHigh  : LREAL := 5.0;             (* 电流偏高置位线，[A]，须 > 0 / the high current set point *)
    fCurrHyst  : LREAL := 0.5;             (* 电流回差，[A]，域 [0, fCurrHigh) / the current hysteresis *)
    tNoPart    : TIME := T#10S;            (* 无件确认延时，[ms] / the no-part confirmation delay *)
    tConfirm   : TIME := T#5S;             (* 电流确认延时，[ms] / the current confirmation delay *)
END_VAR
VAR_OUTPUT
    bJam       : BOOL;                     (* 堵料判定（保持型，复位解除），[标志] / the jam verdict, held until reset *)
    bNoPartOk  : BOOL;                     (* 无件判据已确认，[标志] / the no-part criterion confirmed *)
    bHighCurrOk : BOOL;                    (* 电流判据已确认，[标志] / the high current criterion confirmed *)
    bBusy      : BOOL;                     (* 任一侧确认计时进行中，[标志] / either confirmation timer is running *)
    bValid     : BOOL;                     (* 出口可信（无锁存故障），[标志] / the outlets are trustworthy *)
    bError     : BOOL;                     (* 故障标志（含堵料判定），[标志] / the fault flag, the jam included *)
    nErrCode   : UDINT;                    (* 错误码，0 = 正常，锁存回放 / the error id, 0 = ok, replayed *)
END_VAR
VAR
    _rtReset    : R_TRIG;                  (* 复位上升沿实例（无条件调用）/ the reset rising edge instance *)
    _tonNoPart  : TON;                     (* 无件确认延时实例（无条件调用）/ the no-part confirmation timer *)
    _tonConfirm : TON;                     (* 电流确认延时实例（无条件调用）/ the current confirmation timer *)
    _bJam       : BOOL;                    (* 堵料保持量，仅 bReset 上升沿解除 / the held jam bit *)
    _bFault     : BOOL;                    (* 组态 / 输入故障锁存位 / the configuration and input fault latch *)
    _nCodeLatch : UDINT;                   (* 故障锁存码（0601 / 0602）/ the fault code latch *)
    _bCfgBad    : BOOL;                    (* 组态非法标志（逐拍重算）/ the configuration fault flag *)
    _bInBad     : BOOL;                    (* 电流非有限标志（逐拍重算）/ the current fault flag *)
    _bNoPartCond : BOOL;                   (* 无件条件（含自保持与运行前置），[标志] / the no-part condition *)
    _bCurrCond  : BOOL;                    (* 电流条件（含自保持与回差），[标志] / the current condition *)
END_VAR
VAR CONSTANT
    DL_CJD_FMAX : LREAL := 1.0E30;         (* 非有限筛查幅值上限，[A] / the finiteness screening cap *)
END_VAR

// 段 1｜出口预置（R256 统一出口预置）/ segment 1, preset every outlet
bJam        := FALSE;                      // 堵料判定预清零（真值在段 9 由保持量映射）/ preset the jam verdict false
bNoPartOk   := FALSE;                      // 无件确认位预清零 / preset the no-part flag false
bHighCurrOk := FALSE;                      // 电流确认位预清零 / preset the high current flag false
bBusy       := FALSE;                      // 忙碌标志预清零 / preset the busy flag false
bValid      := FALSE;                      // 可用标志预置假，健康路径再置真 / preset valid false
bError      := FALSE;                      // 故障标志预清零 / preset the error flag false
nErrCode    := 0;                          // 错误码预置无错 / preset the code to zero
_bNoPartCond := FALSE;                     // 无件条件预清零 / preset the no-part condition false
_bCurrCond   := FALSE;                     // 电流条件预清零 / preset the current condition false

// 段 2｜沿检测与定时器无条件调用（规则 ⑦）/ segment 2, the reset edge instance
_rtReset(CLK := bReset);                   // 复位沿，每周期无条件刷新 / the reset edge, refreshed every scan

// 段 3｜堵料解除：唯一可到达的清除边（R188）/ segment 3, the only jam release edge
IF _rtReset.Q THEN                         // 复位上升沿 / the reset rising edge
    _bJam := FALSE;                        // 解除堵料保持 / release the jam hold
END_IF

// 段 4｜组态守卫（R272 逐项点名）/ segment 4, the configuration guard
_bCfgBad := (fCurrHigh <= 0.0)                                       // 置位线非正 / a non positive set point
         OR (fCurrHyst < 0.0)                                        // 回差为负 / a negative hysteresis
         OR (fCurrHyst >= fCurrHigh)                                 // 回差吞没置位线（释放线为负，判据恒自保持）/ the hysteresis swallows the set point
         OR (fCurrHigh <> fCurrHigh) OR ((fCurrHigh - fCurrHigh) <> 0.0) OR (ABS(fCurrHigh) > DL_CJD_FMAX)
         OR (fCurrHyst <> fCurrHyst) OR ((fCurrHyst - fCurrHyst) <> 0.0) OR (ABS(fCurrHyst) > DL_CJD_FMAX);

// 段 5｜输入守卫：电机电流非有限 / segment 5, the current input guard
_bInBad := (fMotorA <> fMotorA) OR ((fMotorA - fMotorA) <> 0.0) OR (ABS(fMotorA) > DL_CJD_FMAX);

// 段 6｜首次成因锁存（故障期不重推断，R189）/ segment 6, the first cause latch
IF NOT _bFault THEN                        // 未锁存才登记 / register only while healthy
    IF _bCfgBad THEN                       // 组态非法优先 / the configuration first
        _bFault     := TRUE;               // 置锁存 / latch it
        _nCodeLatch := 16#0002_0601;       // 故障级：组态非法 / fault level: an illegal configuration
    ELSIF _bInBad THEN                     // 电流非有限 / the current is non finite
        _bFault     := TRUE;               // 置锁存 / latch it
        _nCodeLatch := 16#0002_0602;       // 故障级：输入非有限 / fault level: an input is non finite
    END_IF
END_IF

// 段 7｜两侧判据条件（含自保持与回差，IN 用显式条件）/ segment 7, both criterion conditions
IF bEn AND NOT _bFault THEN                // 使能且无故障才评估条件 / evaluate only while enabled and healthy
    _bNoPartCond := bConvRun AND (NOT bDownPart OR _tonNoPart.Q);                       // 无件条件：运行中且无件（确认后自保持到有件）
    _bCurrCond   := bConvRun AND ((fMotorA > fCurrHigh) OR (_tonConfirm.Q AND (fMotorA > (fCurrHigh - fCurrHyst)))); // 电流条件：超置位线或已确认且未破回差线
ELSE                                       // 失能或故障 / disabled or faulted
    _bNoPartCond := FALSE;                 // 条件清零，计时器随之复位 / clear the condition, the timer resets
    _bCurrCond   := FALSE;                 // 条件清零 / clear the condition
END_IF

// 段 8｜定时器无条件周期调用（规则 ⑦）/ segment 8, unconditional timer calls
_tonNoPart(IN := _bNoPartCond, PT := tNoPart);     // 无件确认计时，每周期无条件刷新 / the no-part timer
_tonConfirm(IN := _bCurrCond, PT := tConfirm);     // 电流确认计时，每周期无条件刷新 / the current timer

// 段 9｜确认位与堵料合成（判据合成点在定时器之后，本拍即可观测）/ segment 9, the synthesis
bNoPartOk   := bEn AND NOT _bFault AND _tonNoPart.Q;    // 无件判据确认 / the no-part criterion confirmed
bHighCurrOk := bEn AND NOT _bFault AND _tonConfirm.Q;   // 电流判据确认 / the current criterion confirmed
bBusy       := bEn AND NOT _bFault AND ((_bNoPartCond AND NOT _tonNoPart.Q) OR (_bCurrCond AND NOT _tonConfirm.Q)); // 任一侧计时中
IF bNoPartOk AND bHighCurrOk THEN          // 双判据同时确认 / both criteria confirmed together
    _bJam := TRUE;                         // 置堵料保持量（锁存至复位）/ hold the jam until a reset
END_IF

// 段 10｜出口映射（名实双出口同源，R191；故障码优先级写入）/ segment 10, the outlet mapping
bJam     := _bJam;                         // 堵料判定出口 = 保持量 / the jam outlet mirrors the hold
bError   := _bJam OR _bFault;              // 故障标志 = 堵料 或 锁存故障 / the fault flag, the jam or the latch
bValid   := bEn AND NOT _bJam AND NOT _bFault; // 出口可信条件 / the outlets are trustworthy
IF _bJam THEN                              // 堵料优先归因（过程故障优先于组态）/ the jam takes precedence
    nErrCode := 16#0002_0603;              // 故障级：堵料 / fault level: a jam was detected
ELSE                                       // 非堵料 / no jam
    nErrCode := _nCodeLatch;               // 回放组态 / 输入锁存码 / replay the configuration or input code
END_IF
END_FUNCTION_BLOCK

(* ---- FB_DL_ConveyorSlipWatch.st ---- *)
(*
  Name        : FB_DL_ConveyorSlipWatch
  Category    : DL_Device
  Version     : 1.0.0
  Purpose     : 输送带打滑检测：带速与驱动辊线速差折算打滑率，叠加电流负载判据（轻载不判滑），超限经确认延时锁存报警；/ Conveyor slip watch: slip ratio from belt vs drive-roll surface speed, gated by a current load criterion, confirmed then latched over the threshold
  溯源        : 借 t2-2-lbp 的分类/参数域组织，clean-room 实现
  Boundary    : ① 组态闸：速度下限/打滑率上限/电流下限/确认延时任一越域 → 锁存故障；
                ② 除零前置：打滑率除子取驱动辊速绝对值，须 >= 速度下限（组态闸保证）才计算；
                ③ 非有限速度/电流该拍不判（保留上拍结果，防污染判据）；
                ④ 确认延时 TON 串 eMon 相位闸（族③：eIdle/eFault 不计时），段 0 无 IF 包裹；
                ⑤ 负打滑（带速 > 辊速，属测量倒置）不判滑但置诊断位 bRatioInvert；
                ⑥ 本件为诊断层，不停机（属主边界）。
*)
TYPE E_DL_CswState :
(
    eIdle  := 0,                             (* 未使能 / Disabled *)
    eMon   := 10,                            (* 打滑监视运行 / Monitoring *)
    eFault := 90                             (* 故障锁存相 / Fault latched *)
);
END_TYPE

TYPE E_DL_CswCause :
(
    eNone       := 0,                        (* 无故障成因 / No cause *)
    eCfgIllegal := 1,                        (* 组态非法：速度/比率/电流/延时越域 / Illegal config *)
    eSlip       := 2,                        (* 打滑确认（带速滞后辊速） / Confirmed slip *)
    ePhaseBad   := 3                         (* 非法相位兜底 / Illegal phase fallback *)
);
END_TYPE

FUNCTION_BLOCK FB_DL_ConveyorSlipWatch
VAR_INPUT
    fBeltSpeed  : REAL := 0.0;               (* 带速实测（带秤/编码器折算）[m/s] / Measured belt speed *)
    fRollSpeed  : REAL := 0.0;               (* 驱动辊线速度实测 [m/s] / Drive-roll surface speed *)
    fSpdMin     : REAL := 0.2;               (* 速度计算下限（除子域 + 运行判定），域 > 0 [m/s] / Speed floor for divisor and run gating *)
    fSlipMax    : REAL := 5.0;               (* 打滑率报警上限，域 > 0 [%] / Slip ratio limit, > 0 *)
    fCurrent    : REAL := 0.0;               (* 驱动电机电流实测 [A] / Drive motor current *)
    fCurrentMin : REAL := 2.0;               (* 负载电流下限（轻载不判滑），域 > 0 [A] / Load current floor *)
    tConfirm    : TIME := T#2S;              (* 打滑确认延时，域 > T#0S [ms] / Slip confirm delay, > 0 *)
    bRunning    : BOOL := FALSE;             (* 输送机运行命令电平 [-] / Conveyor run command *)
    bEnable     : BOOL := TRUE;              (* 监视使能 [-] / Enable *)
    bReset      : BOOL := FALSE;             (* 复位命令，上升沿清报警与故障 [-] / Reset command *)
END_VAR
VAR_OUTPUT
    fSlipRatio  : REAL;                      (* 打滑率（实时派生，速度不足时为 0）[%] / Slip ratio *)
    bLoaded     : BOOL;                      (* 负载在位（电流 >= 下限）[-] / Load present *)
    bRatioInvert: BOOL;                      (* 打滑率为负（测量倒置诊断位）[-] / Negative slip ratio diagnostic *)
    bSlip       : BOOL;                      (* 打滑报警锁存（复位沿清）[-] / Slip alarm latched *)
    eState      : E_DL_CswState;             (* 状态出口 / State outlet *)
    eCause      : E_DL_CswCause;             (* 故障成因出口（R190 归因唯一） / Fault cause outlet *)
    bError      : BOOL;                      (* 故障锁存标志 [-] / Fault latch flag *)
END_VAR
VAR
    _eState  : E_DL_CswState := E_DL_CswState.eIdle;     (* 内部相位（CASE 唯一写入目标） / Internal phase *)
    _eCause  : E_DL_CswCause := E_DL_CswCause.eNone;     (* 故障成因锁存量 / Latched cause *)
    rtReset  : R_TRIG;                       (* 复位沿实例，段 0 无条件调用 / Reset edge instance *)
    tonConf  : TON;                          (* 打滑确认延时计时器（IN 由判据派生 + 相位闸） / Slip confirm timer *)
    _bFault  : BOOL;                         (* 故障锁存位 / Latched fault bit *)
    _bCfgBad : BOOL;                         (* 组态非法当拍量 / Illegal config this scan *)
    _bFin    : BOOL;                         (* 输入有限性当拍量（三输入联合） / Input finiteness joint *)
    _bRun    : BOOL;                         (* 速度达标运行当拍量（两速度均 >= 下限） / Speeds above floor *)
    _bLoad   : BOOL;                         (* 负载在位当拍量 / Load present this scan *)
    _fRatio  : REAL;                         (* 打滑率中间量 [%] / Slip ratio intermediate *)
    _bSlipRaw: BOOL;                         (* 打滑原始判据当拍量 / Raw slip verdict *)
END_VAR
VAR CONSTANT
    DL_CSW_EPS    : REAL := 1.0E-6;          (* 判零容差 [-] / Epsilon *)
    DL_CSW_HUND   : REAL := 100.0;           (* 百分数换算常量（乘性常量）[-] / Percent scale constant *)
END_VAR

(* —— 段 0：当拍判据派生 + 实例无条件刷新（R228A；R_TRIG/TON 全在段 0，无 IF 包裹） —— *)
_bCfgBad := (fSpdMin <= DL_CSW_EPS)                                            (* 速度下限正域闸（兼除子域闸） / Speed floor gate *)
            OR (fSlipMax <= DL_CSW_EPS)                                        (* 打滑率上限正域闸 / Slip limit gate *)
            OR (fCurrentMin <= DL_CSW_EPS)                                     (* 电流下限正域闸 / Current floor gate *)
            OR NOT (tConfirm > T#0S);                                          (* 确认延时正域闸 / Confirm delay gate *)
rtReset(CLK := bReset);                                                        (* 复位沿每拍必调 / Reset edge every scan *)
_bFin := (fBeltSpeed = fBeltSpeed) AND (fRollSpeed = fRollSpeed)               (* 速度 NaN 自反闸 / Speeds NaN gates *)
            AND (fCurrent = fCurrent)                                          (* 电流 NaN 自反闸 / Current NaN gate *)
            AND ((fBeltSpeed - fBeltSpeed) = (fBeltSpeed - fBeltSpeed))        (* 带速 Inf 差判闸 / Belt speed Inf gate *)
            AND ((fRollSpeed - fRollSpeed) = (fRollSpeed - fRollSpeed))        (* 辊速 Inf 差判闸 / Roll speed Inf gate *)
            AND ((fCurrent - fCurrent) = (fCurrent - fCurrent));               (* 电流 Inf 差判闸 / Current Inf gate *)
_bRun := _bFin AND (ABS(fRollSpeed) >= fSpdMin) AND (ABS(fBeltSpeed) >= fSpdMin);   (* 两速度均达下限才计算比率（除子域闸边界②） / Both speeds above floor *)
_fRatio := 0.0;                                                                (* 打滑率中间量预置（速度不足时保持 0，出口确定值） / Ratio preset zero *)
IF _bRun THEN
    _fRatio := (fRollSpeed - fBeltSpeed) / ABS(fRollSpeed) * DL_CSW_HUND;      (* 打滑率 = (辊速-带速)/|辊速|：除子 |辊速| >= 下限已闸 [%] / Slip ratio, divisor gated *)
END_IF
_bLoad := _bFin AND (fCurrent >= fCurrentMin);                                 (* 负载在位：电流达下限 / Load present *)
_bSlipRaw := _bFin AND _bRun AND _bLoad AND (_fRatio > fSlipMax);              (* 原始判据：运行 + 负载 + 超限（三者同证） / Raw slip verdict *)
tonConf(IN := (_eState = E_DL_CswState.eMon) AND bRunning AND _bSlipRaw, PT := tConfirm);   (* 确认延时：判据持续才计时，串 eMon 相位闸 / Confirm timer with phase gate *)

(* —— 段 1：单拍量预清零（R107） —— *)
bLoaded := FALSE;                                                              (* 负载指示预清 / Load preset *)
bRatioInvert := FALSE;                                                         (* 倒置诊断位预清 / Invert preset *)
fSlipRatio := 0.0;                                                             (* 打滑率出口预清 / Ratio outlet preset *)

(* —— 段 2：复位沿处理（作用域：清故障 + 清报警 + 迁 eIdle，R283 逐项声明） —— *)
IF rtReset.Q THEN
    _bFault := FALSE;                                                          (* 清故障锁存 / Clear fault *)
    _eCause := E_DL_CswCause.eNone;                                            (* 清成因 / Clear cause *)
    bSlip := FALSE;                                                            (* 清打滑报警锁存 / Clear slip latch *)
    _eState := E_DL_CswState.eIdle;                                            (* 迁未使能相 / Back to idle *)
END_IF

(* —— 段 3：组态故障锁存（锁存至复位沿，R189） —— *)
IF _bCfgBad AND NOT _bFault THEN
    _bFault := TRUE;                                                           (* 锁存故障位 / Latch fault *)
    _eCause := E_DL_CswCause.eCfgIllegal;                                      (* 成因：组态非法 / Cause: illegal config *)
    _eState := E_DL_CswState.eFault;                                           (* 同步迁故障相 / Migrate to fault *)
END_IF

(* —— 段 4：CASE 主状态机（ELSE 兜底迁 eFault，红线 6） —— *)
CASE _eState OF
    E_DL_CswState.eIdle:                                                       (* 未使能：出口确定值 / Disabled *)
        fSlipRatio := 0.0;                                                     (* 失能清打滑率出口 / Clear ratio outlet *)
        bSlip := FALSE;                                                        (* 失能清报警出口 / Clear slip outlet *)
        bLoaded := FALSE;                                                      (* 失能清负载出口 / Clear load outlet *)
        bRatioInvert := FALSE;                                                 (* 失能清倒置出口 / Clear invert outlet *)
        IF bEnable AND NOT _bFault THEN
            _eState := E_DL_CswState.eMon;                                     (* 使能进入监视 / Enter monitoring *)
        END_IF
    E_DL_CswState.eMon:                                                        (* 监视相：比率派生 + 确认锁存 / Monitoring *)
        IF NOT bEnable THEN
            _eState := E_DL_CswState.eIdle;                                    (* 失能回未使能 / Back to idle *)
        ELSE
            fSlipRatio := _fRatio;                                             (* 打滑率出口（实时派生，R191） / Ratio outlet *)
            bLoaded := _bLoad;                                                 (* 负载出口（名实同源） / Load outlet *)
            bRatioInvert := _bFin AND _bRun AND (_fRatio < 0.0);               (* 负比率诊断：带速 > 辊速（测量倒置） / Inverted ratio diagnostic *)
            IF tonConf.Q THEN                                                  (* 判据持续满确认延时：锁存报警 / Confirm elapsed: latch alarm *)
                bSlip := TRUE;                                                 (* 打滑报警锁存（复位沿清） / Latch slip *)
                _bFault := TRUE;                                               (* 同步故障锁存（R45 配对） / Latch fault *)
                _eCause := E_DL_CswCause.eSlip;                                (* 成因：打滑 / Cause: slip *)
            END_IF
        END_IF
    E_DL_CswState.eFault:                                                      (* 故障相：冻结保持末值，仅复位沿出 / Fault *)
        ;                                                                      (* 锁存回放（R28） / Replay from latch *)
    ELSE                                                                       (* 非法相位兜底迁安全态 / Illegal phase fallback *)
        _eState := E_DL_CswState.eFault;                                       (* 迁故障相 / To fault *)
        _bFault := TRUE;                                                       (* 同步锁存 / Latch *)
        _eCause := E_DL_CswCause.ePhaseBad;                                    (* 成因：非法相位 / Cause: illegal phase *)
END_CASE

(* —— 段 5：出口映射（bError/eState 同源，R191） —— *)
bError := _bFault;                                                             (* 故障标志镜像 / Fault flag mirror *)
eState := _eState;                                                             (* 状态出口 / State outlet *)
eCause := _eCause;                                                             (* 成因出口 / Cause outlet *)
END_FUNCTION_BLOCK

(* ---- FB_DL_CoolantFlowAudit.st ---- *)
// =====================================================================
// FB_DL_CoolantFlowAudit.st
// 机台冷却水多支路流量审计（欠流确认窗 + 迟滞锁存 + 首出三律定位）
// Multi-branch coolant flow audit with underflow confirm and first-out
// 所属子库: DL_Device    版本: v1.0.0    兼容: CODESYS V3.5+ / TwinCAT 3 / 汇川 InoProShop
// 码位: 16#0003_03E3 ~ 16#0003_03E7 (本件独占 5 槽, 勿复用)
// 溯源: 道莅 clean-room 防御性实现
//       来源组标签: semiconductor, coolant, flow-audit, alarm-management
// 修改记录: R30 初版 (ROUND_PLAN_R30 序 3)
// =====================================================================
FUNCTION_BLOCK FB_DL_CoolantFlowAudit
VAR_INPUT
    bEnable       : BOOL  := FALSE;   // 使能 / Enable
    afFlow_Lpm    : ARRAY[1..8] OF REAL;   // 各支路流量 0~500 L/min / Branch flow [L/min]
    afMinFlow_Lpm : ARRAY[1..8] OF REAL;   // 各支路欠流阈值 0~500 L/min / Branch underflow threshold [L/min]
    tConfirm      : TIME  := T#2S;    // 欠流确认窗 T#10MS~T#60S / Underflow confirm window [s]
    fHyst_Lpm     : REAL  := 2.0;     // 欠流解除迟滞 0~50 L/min / Release hysteresis [L/min]
END_VAR
VAR_OUTPUT
    uwUnderMask   : WORD  := 0;       // 欠流位掩码, 位 0..7 对应支路 1..8 / Underflow mask, bit0..7 = branch 1..8
    uFirstOut     : USINT := 0;       // 首出支路号 1~8, 0 = 无 / First-out branch, 0 = none
    bAllOk        : BOOL  := FALSE;   // 全部支路正常 / All branches ok
    eErr          : UDINT := 16#0003_03E3;  // 错误码 / Error code
END_VAR
VAR
    aTonConf      : ARRAY[1..8] OF TON;   // 各支路欠流确认定时器, 每拍无条件刷新 / Per-branch confirm timers, refreshed every cycle
    abUnderLatch  : ARRAY[1..8] OF BOOL;  // 各支路欠流锁存 / Per-branch underflow latch
    abSensorFlt   : ARRAY[1..8] OF BOOL;  // 各支路传感器故障标记 / Per-branch sensor fault flag
    bCfgErr       : BOOL  := FALSE;   // 组态非法标记 / Configuration error flag
    bSnsErr       : BOOL  := FALSE;   // 任一支路传感器故障标记 / Any-branch sensor fault flag
    uFirstLatch   : USINT := 0;       // 首出锁存支路号 / First-out latched branch
    uZi           : INT   := 1;       // 1..8 数组下标 / Array subscript 1..8
END_VAR

// ---------------------------------------------------------------------
// 代码位表（本件独占, 勿复用）:
//   16#0003_03E3 信息 全部支路正常
//   16#0003_03E4 故障 组态非法（欠流阈值或迟滞非有限, 或越出 0~500/0~50 L/min 合法域）
//   16#0003_03E5 故障 任一支路流量非有限/为负/超量程（传感器故障, 独立于欠流判据）
//   16#0003_03E6 故障 存在确认欠流支路（掩码非零）, 解除式 = 对应支路流量恢复到阈值+迟滞以上
//   16#0003_03E7 信息 待机未使能
// ---------------------------------------------------------------------

// ---- 守卫闸: 迟滞与逐支路阈值合法域 / Gate: hysteresis and per-branch threshold validity ----
bCfgErr := FALSE;               // 组态错误标记复位 / Reset config error flag
IF (fHyst_Lpm <> fHyst_Lpm) OR (fHyst_Lpm < 0.0) OR (fHyst_Lpm > 50.0) THEN
    bCfgErr := TRUE;            // 迟滞非法 / Illegal hysteresis
END_IF
IF NOT bCfgErr THEN
    FOR uZi := 1 TO 8 DO
        IF (afMinFlow_Lpm[uZi] <> afMinFlow_Lpm[uZi])
           OR (afMinFlow_Lpm[uZi] < 0.0) OR (afMinFlow_Lpm[uZi] > 500.0) THEN
            bCfgErr := TRUE;    // 阈值越界即组态故障 / Threshold out of domain = config fault
        END_IF
    END_FOR
END_IF

// ---- 逐支路传感器故障判: 非有限/负值/超量程, 独立于欠流判据 / Per-branch sensor fault judge ----
bSnsErr := FALSE;               // 传感器故障标记复位 / Reset sensor fault flag
FOR uZi := 1 TO 8 DO
    abSensorFlt[uZi] := (afFlow_Lpm[uZi] <> afFlow_Lpm[uZi])
                     OR (afFlow_Lpm[uZi] < 0.0)
                     OR (afFlow_Lpm[uZi] > 500.0);  // 非有限自反判或越域 / Non-finite or out of domain
    IF abSensorFlt[uZi] THEN
        bSnsErr := TRUE;        // 置总传感器故障标记 / Set overall sensor fault flag
    END_IF
END_FOR

// ---- 欠流确认定时器无条件周期刷新 + 锁存/解除 / Confirm timers unconditional refresh, latch and release ----
FOR uZi := 1 TO 8 DO
    IF bEnable AND (NOT bCfgErr) AND (NOT abSensorFlt[uZi]) AND (NOT abUnderLatch[uZi]) THEN
        // 进入条件: 流量低于阈值计时, 窗内瞬时恢复自动清零计时（抖动不误报）
        // Enter: below threshold timing; transient recovery resets timing in window
        aTonConf[uZi](IN := afFlow_Lpm[uZi] < afMinFlow_Lpm[uZi], PT := tConfirm);
        IF aTonConf[uZi].Q AND (afFlow_Lpm[uZi] < afMinFlow_Lpm[uZi]) THEN
            abUnderLatch[uZi] := TRUE;      // 确认欠流锁存 / Confirm underflow latch
        END_IF
    ELSE
        aTonConf[uZi](IN := FALSE, PT := tConfirm);     // 非候选支路显式复位 / Explicit reset for non-candidates
    END_IF
    // 解除: 流量恢复到阈值+迟滞以上 / Release: flow above threshold plus hysteresis
    IF abUnderLatch[uZi] AND (NOT abSensorFlt[uZi])
       AND (afFlow_Lpm[uZi] >= (afMinFlow_Lpm[uZi] + fHyst_Lpm)) THEN
        abUnderLatch[uZi] := FALSE;     // 解除欠流锁存 / Release underflow latch
    END_IF
    // 传感器故障拍欠流判据失效, 强制解除该支路锁存 / Sensor fault voids underflow judge
    IF abSensorFlt[uZi] THEN
        abUnderLatch[uZi] := FALSE;     // 强制解除 / Forced release
    END_IF
END_FOR

// ---- 欠流位掩码汇总 / Underflow mask aggregation ----
uwUnderMask := 0;                   // 掩码复位 / Reset mask
FOR uZi := 1 TO 8 DO
    IF abUnderLatch[uZi] THEN
        uwUnderMask := uwUnderMask OR SHL(WORD#1, uZi - 1);     // 移位量 0..7 小于字宽, 合规 / Shift 0..7 within word width
    END_IF
END_FOR

// ---- 首出三律: 未锁存才仲裁, 同拍取最小支路号, 解除在仲裁后（掩码全清时释放）
//      First-out laws: arbitrate only if not latched, min branch per cycle, release after mask clears ----
IF (uFirstLatch = 0) AND (uwUnderMask <> 0) THEN
    FOR uZi := 1 TO 8 DO
        IF (uFirstLatch = 0) AND abUnderLatch[uZi] THEN
            uFirstLatch := INT_TO_USINT(uZi);   // 升序扫描, 首个命中即最小支路号 / Ascending scan picks min branch
        END_IF
    END_FOR
END_IF
IF uwUnderMask = 0 THEN
    uFirstLatch := 0;               // 全部支路恢复后释放首出锁存 / Release first-out when all clear
END_IF
uFirstOut := uFirstLatch;           // 输出首出支路号 / Output first-out branch

// ---- 全正常输出 / All-ok output ----
bAllOk := bEnable AND (NOT bCfgErr) AND (NOT bSnsErr) AND (uwUnderMask = 0);

// ---- 错误码仲裁（每拍重算, 故障解除可达）/ Error arbitration, releasable ----
IF bCfgErr THEN
    eErr := 16#0003_03E4;           // 组态非法 / Configuration fault
ELSIF bSnsErr THEN
    eErr := 16#0003_03E5;           // 传感器故障 / Sensor fault
ELSIF uwUnderMask <> 0 THEN
    eErr := 16#0003_03E6;           // 存在欠流支路 / Underflow present
ELSIF NOT bEnable THEN
    eErr := 16#0003_03E7;           // 待机未使能 / Standby
ELSE
    eErr := 16#0003_03E3;           // 全部正常 / All normal
END_IF

END_FUNCTION_BLOCK

(* ---- FB_DL_CoolantLoopBal.st ---- *)
// =====================================================================
// FB_DL_CoolantLoopBal.st
// 机台冷却水 4 支路流量均衡（增量总和强制归零，保总流量守恒）
// Coolant 4-branch flow balance FB
// 码位: 16#0003_03C0 ~ 16#0003_03C4 (本件独占 5 槽)
// 修改记录: R29 初版 (按 DISPATCH_R29 序 7)
// =====================================================================
FUNCTION_BLOCK FB_DL_CoolantLoopBal
VAR_INPUT
    bEnable       : BOOL  := FALSE;    // 使能 / Enable
    abFlowValid   : ARRAY[1..4] OF BOOL;   // 支路流量有效 / Branch flow valid
    afFlow_lpm    : ARRAY[1..4] OF REAL;   // 支路流量 0~500 L/min / Branch flow [L/min]
    fFlowMin_lpm  : REAL  := 5.0;      // 均衡投入最低总流量 >0 L/min / Min total flow [L/min]
    fGain         : REAL  := 0.5;      // 均衡增益 0.05~2.0 / Balance gain [-]
    fTrimMax_pct  : REAL  := 5.0;      // 单拍最大阀位增量 0.1~20 % / Max step [%]
    fDevMax_pct   : REAL  := 20.0;     // 失衡报警阈值 1~100 % / Imbalance alarm [%]
    tWin          : TIME  := T#2S;     // 均值窗口 T#200MS~T#30S / Averaging window [s]
END_VAR
VAR_OUTPUT
    afValve_pct   : ARRAY[1..4] OF REAL;    // 支路阀位 0~100 %（本件独占写）/ Branch valve [%]
    fFlowAvg_lpm  : REAL;               // 窗口平均总流量 L/min / Average total flow [L/min]
    fImb_pct      : REAL;               // 最大支路偏差 % / Max imbalance [%]
    bBalanced     : BOOL;               // 失衡 ≤ 5 % / Balanced
    bFrozen       : BOOL;               // 冻结中 / Frozen
    eErr          : UDINT;              // 错误码 / Error code
END_VAR
VAR
    aDelta        : ARRAY[1..4] OF REAL;    // 各路增量暂存 / Per-branch delta [%]
    fDeltaSum     : REAL;               // 增量代数和 / Delta sum [%]
    fDeltaMean    : REAL;               // 增量均值 / Delta mean [%]
    uValidCnt     : UDINT;              // 有效支路数 / Valid branch count
    uIdx          : UDINT;              // 循环下标 / Loop index
    uZi           : INT;                // 1..4 数组下标 / Array subscript 1..4
    fTotal        : REAL;               // 有效支路总流量 / Total valid flow [L/min]
    fAvgBranch    : REAL;               // 有效支路平均流量 / Average branch flow [L/min]
    fImbMax       : REAL;               // 最大偏差 / Max imbalance [%]
    fDevRel       : REAL;               // 支路相对偏差 / Relative deviation [-]
    tWinS         : REAL;               // 窗口秒值 / Window in seconds [s]
    fBase         : REAL;               // 均值窗口基准（首拍锁定）/ Window baseline, locked on first cycle [L/min]
    xHasBase      : BOOL  := FALSE;     // 基准已锁定标记 / Baseline locked flag
    xFirstScan    : BOOL  := TRUE;      // 首扫标记 / First-scan flag
END_VAR

// ---------------------------------------------------------------------
// 代码位表（本件独占，勿复用）:
//   16#0003_03C0 信息 均衡运行正常
//   16#0003_03C1 故障 流量值非有限 / tWin 非法
//   16#0003_03C2 故障 fGain ≤ 0 / fTrimMax_pct ≤ 0 / fFlowMin_lpm ≤ 0（组态错）
//   16#0003_03C3 信息 单支路阀位触 0/100 % 或流量计无效 → 该路冻结；有效支路 < 2 → 不均衡
//   16#0003_03C4 信息 总流量 < fFlowMin_lpm → 全冻结（bFrozen=TRUE），fImb_pct 照算供上位看
// ---------------------------------------------------------------------

// ---- 窗口转秒 / Window to seconds ----
tWinS := TIME_TO_REAL(tWin) / 1000.0;       // 秒值 / Seconds [s]

// ---- 非有限与窗口合法性闸 / Finite and window validity gate ----
IF (tWin = T#0MS) OR (tWinS < 0.2) OR (tWinS > 30.0)
   OR (fGain <> fGain) OR (ABS(fGain) >= 1.0E12)
   OR (fFlowMin_lpm <> fFlowMin_lpm) OR (ABS(fFlowMin_lpm) >= 1.0E12)
   OR (fTrimMax_pct <> fTrimMax_pct) OR (ABS(fTrimMax_pct) >= 1.0E12) THEN
    bFrozen := TRUE;            // 安全冻结 / Safe freeze
    eErr    := 16#0003_03C1;    // 故障码 / Fault code
    RETURN;                     // 阀位保持不动 / Valves hold
END_IF

// ---- 逐支路流量非有限判界（多 ARRAY 各自判）/ Per-branch finite check ----
FOR uZi := 1 TO 4 DO
    IF (afFlow_lpm[uZi] <> afFlow_lpm[uZi]) OR (ABS(afFlow_lpm[uZi]) >= 1.0E12) THEN
        bFrozen := TRUE;        // 安全冻结 / Safe freeze
        eErr    := 16#0003_03C1;    // 故障码 / Fault code
        RETURN;                 // 阀位保持不动 / Valves hold
    END_IF
END_FOR

// ---- 组态错闸 / Configuration fault gate ----
IF (fGain <= 0.0) OR (fTrimMax_pct <= 0.0) OR (fFlowMin_lpm <= 0.0) THEN
    bFrozen := TRUE;            // 安全冻结 / Safe freeze
    eErr    := 16#0003_03C2;    // 故障码 / Fault code
    RETURN;                     // 本拍结束 / End of cycle
END_IF

// ---- 首扫初始化：阀位从外部给定基准起（R16 首扫纪律）/ First-scan init ----
IF xFirstScan THEN
    FOR uZi := 1 TO 4 DO
        afValve_pct[uZi] := 50.0;   // 阀位初值 50 % / Valve init 50 %
        aDelta[uZi] := 0.0;     // 增量清零 / Delta cleared
    END_FOR
    xFirstScan := FALSE;        // 清标记 / Clear flag
END_IF

// ---- 使能撤销：全冻结（阀位保持）/ Disable: hold valves ----
IF NOT bEnable THEN
    bFrozen   := FALSE;         // 非欠流冻结 / Not underflow freeze
    bBalanced := FALSE;         // 结论失效 / Verdict invalid
    eErr      := 16#0003_03C0;  // 信息级：空闲 / Info: idle
    RETURN;                     // 阀位保持不动 / Valves hold
END_IF

// ---- 有效支路统计 / Valid branch counting ----
uValidCnt := 0;                 // 计数清零 / Reset count
fTotal := 0.0;                  // 总量清零 / Reset total
FOR uZi := 1 TO 4 DO
    IF abFlowValid[uZi] THEN
        uValidCnt := uValidCnt + 1;     // 有效计数 / Count valid
        fTotal := fTotal + afFlow_lpm[uZi]; // 累加流量 / Accumulate flow
    END_IF
END_FOR

// ---- 均值分母钳 ≥1 / Denominator clamp ≥1 ----
IF uValidCnt >= 1 THEN
    fAvgBranch := fTotal / UDINT_TO_REAL(uValidCnt);    // 平均支路流量 / Average branch flow
ELSE
    fAvgBranch := 0.0;          // 无有效路 / No valid branch
END_IF
fFlowAvg_lpm := fAvgBranch * UDINT_TO_REAL(uValidCnt);  // 窗口平均总流量（有效口径）/ Average total flow

// ---- 有效支路数 < 2 → 不均衡并置槽 4（单支路无相对量）/ Fewer than 2 valid branches ----
IF uValidCnt < 2 THEN
    bFrozen := TRUE;            // 冻结 / Freeze
    bBalanced := FALSE;         // 结论失效 / Verdict invalid
    fImb_pct := 0.0;            // 偏差无意义置 0 / Imbalance meaningless
    eErr := 16#0003_03C3;       // 信息级：路数不足 / Info: insufficient branches
    RETURN;                     // 阀位保持不动 / Valves hold
END_IF

// ---- 失衡统计（照算供上位看）/ Imbalance statistics (always computed) ----
fImbMax := 0.0;                 // 最大偏差复位 / Reset max
FOR uZi := 1 TO 4 DO
    IF abFlowValid[uZi] THEN
        IF fAvgBranch > 0.0 THEN
            fDevRel := ABS(afFlow_lpm[uZi] - fAvgBranch) / fAvgBranch * 100.0;  // 相对偏差 % / Relative deviation [%]
        ELSE
            fDevRel := 0.0;     // 分母保护 / Denominator guard
        END_IF
        IF fDevRel > fImbMax THEN
            fImbMax := fDevRel; // 取最大 / Keep max
        END_IF
    END_IF
END_FOR
fImb_pct := fImbMax;            // 输出最大偏差 / Output max imbalance
bBalanced := (fImbMax <= 5.0);  // 失衡 ≤ 5 % 判 / Balanced verdict

// ---- 总流量欠流 → 全冻结（阀位不变，偏差照算）/ Underflow: freeze all ----
IF fTotal < fFlowMin_lpm THEN
    bFrozen := TRUE;            // 冻结标志 / Frozen flag
    eErr := 16#0003_03C4;       // 信息级：欠流冻结 / Info: underflow freeze
    RETURN;                     // 阀位保持不动 / Valves hold
END_IF
bFrozen := FALSE;               // 正常非冻结 / Not frozen

// ---- 增量计算：先算各路增量再减均值（总和强制归零）/ Deltas then subtract mean ----
FOR uZi := 1 TO 4 DO
    IF abFlowValid[uZi] AND (fAvgBranch > 0.0) THEN
        // 相对偏差 → 阀位增量方向：流量低于均值 → 开阀 / Low flow → open valve
        aDelta[uZi] := fGain * ((fAvgBranch - afFlow_lpm[uZi]) / fAvgBranch) * fTrimMax_pct;    // 原始增量 / Raw delta [%]
    ELSE
        aDelta[uZi] := 0.0;     // 无效路不参与 / Invalid branch excluded
    END_IF
END_FOR
fDeltaSum := 0.0;               // 和清零 / Reset sum
FOR uZi := 1 TO 4 DO
    fDeltaSum := fDeltaSum + aDelta[uZi];   // 代数和 / Algebraic sum
END_FOR
fDeltaMean := fDeltaSum / UDINT_TO_REAL(uValidCnt);     // 增量均值（分母=有效路数）/ Delta mean

// ---- 阀位更新：单拍限幅 + 触限冻结 + 归零修正 / Valve update: slew limit + limit freeze + zero-sum ----
FOR uZi := 1 TO 4 DO
    IF abFlowValid[uZi] THEN
        // 单拍最大增量限幅 / Per-cycle max step clamp
        IF aDelta[uZi] > fTrimMax_pct THEN
            aDelta[uZi] := fTrimMax_pct;    // 正向限幅 / Positive clamp
        ELSIF aDelta[uZi] < -fTrimMax_pct THEN
            aDelta[uZi] := -fTrimMax_pct;   // 负向限幅 / Negative clamp
        END_IF
        // 触限后停止同向修正 / Limit reached: stop same-direction trim
        IF (afValve_pct[uZi] >= 100.0) AND (aDelta[uZi] > 0.0) THEN
            aDelta[uZi] := 0.0;     // 上限同向冻结 / Upper freeze
        ELSIF (afValve_pct[uZi] <= 0.0) AND (aDelta[uZi] < 0.0) THEN
            aDelta[uZi] := 0.0;     // 下限同向冻结 / Lower freeze
        END_IF
    ELSE
        aDelta[uZi] := 0.0;         // 冻结支路增量为 0（不被拉走流量）/ Frozen branch zero delta
    END_IF
END_FOR

// ---- 归零修正重算均值（冻结路不参与均值）/ Re-zero with frozen branches excluded ----
fDeltaSum := 0.0;               // 和清零 / Reset sum
uValidCnt := 0;                 // 计数复位 / Reset count
FOR uZi := 1 TO 4 DO
    IF abFlowValid[uZi] THEN
        fDeltaSum := fDeltaSum + aDelta[uZi];   // 有效路代数和 / Valid sum
        uValidCnt := uValidCnt + 1;     // 有效计数 / Valid count
    END_IF
END_FOR
IF uValidCnt >= 1 THEN
    fDeltaMean := fDeltaSum / UDINT_TO_REAL(uValidCnt);     // 均值 / Mean
ELSE
    fDeltaMean := 0.0;          // 保护 / Guard
END_IF

// ---- 应用增量（减均值保总和守恒）/ Apply deltas minus mean (conservation) ----
FOR uZi := 1 TO 4 DO
    IF abFlowValid[uZi] THEN
        afValve_pct[uZi] := afValve_pct[uZi] + (aDelta[uZi] - fDeltaMean);  // 守恒增量 / Conserved delta
        // 最终阀位钳 0~100 % / Final valve clamp
        IF afValve_pct[uZi] < 0.0 THEN
            afValve_pct[uZi] := 0.0;    // 下限 / Lower clamp
        ELSIF afValve_pct[uZi] > 100.0 THEN
            afValve_pct[uZi] := 100.0;  // 上限 / Upper clamp
        END_IF
    END_IF
END_FOR

// ---- 触限信息级 / At-limit info code ----
FOR uZi := 1 TO 4 DO
    IF abFlowValid[uZi] AND ((afValve_pct[uZi] >= 100.0) OR (afValve_pct[uZi] <= 0.0)) THEN
        eErr := 16#0003_03C3;   // 信息级：触限冻结 / Info: at-limit freeze
        RETURN;                 // 已登记直接返回 / Return after marking
    END_IF
END_FOR

// ---- 正常码 / Normal code ----
eErr := 16#0003_03C0;           // 信息级：均衡正常 / Info: balancing normal

END_FUNCTION_BLOCK

(* ---- FB_DL_CrahGroupEconomizerSeq.st ---- *)
(*
 * FB_DL_CrahGroupEconomizerSeq | C4 | DL_Device
 * 功能：机房群控自然冷却切换序列（机械→过渡→全自然→混合），带焓差滞环与最短驻留       单位：比焓 [kJ/kg]、温度 [℃]、机组数 [台]、rTimeoutS [s]、nFaultCode [INT 码位]
 * 工况边界：判据以户外比焓与回风比焓之差为准（户外 < 回风 − 滞环 → 全自然；|差| ≤ 滞环 → 混合；其余 → 机械）；最短驻留 120 s 由每相 TON 保证，切换只能在驻留满足后进行；nUnitsAvail 须 ≥1，否则 9601；比焓/温度 NaN 或超量程一律 9602/9603 并全回机械侧（安全侧 = 机械冷机）
 * 代数值回代：rOutdoorEnthalpy=45、rReturnEnthalpy=56、hyst=4 → 45 < 52 → 全自然(FREE)；rOutdoor=53 → |53−56|=3 ≤4 → 混合(MIXED)；rOutdoor=60 → 机械(MECH)；nUnitsAvail=0 → 9601（与 spec 判据一致）
 * 开源溯源：clean-room 自研，未复制任何第三方代码（无外部来源）
 *)
(*
 * 码位总账（本件故障码全清单，逐条在实现分支中可到达；故障级锁存回放）：
 * 9601 无可用机组 / 9602 比焓非有限或越量程 / 9603 户外温度非有限或越量程 / 9604 过渡配置非法（rTimeoutS 短于 120 s 最短驻留，自然冷却无法稳定建立）/ 9605 机组数配置越限或状态机兜底（故障锁存，清除沿 = xEnable 下降沿）
 *)

TYPE E_DL_EconMode :
(
    MECH    := 0,       // 全机械制冷，新风阀关闭 | full mechanical cooling, damper closed
    PARTIAL := 10,      // 过渡相，新风阀渐开、机械机组减载 | transition phase, damper ramping open and mechanical units unloading
    FREE    := 20,      // 全自然冷却，新风阀全开、机械全停 | full free cooling, damper fully open and mechanical units off
    MIXED   := 30,      // 混合冷却，新风与机械各半 | mixed cooling, half free and half mechanical
    FAULT   := 90       // 故障相，回机械侧安全值并锁存码位 | fault phase, reverts to the mechanical safe side and latches the code
);
END_TYPE

FUNCTION_BLOCK FB_DL_CrahGroupEconomizerSeq
VAR_INPUT
    xEnable              : BOOL;         // 群控使能（下降沿兼作故障复位沿）| group enable, its falling edge also resets a latched fault
    rOutdoorEnthalpyKJkg : REAL;         // 户外空气比焓 | outdoor air specific enthalpy [kJ/kg]
    rReturnEnthalpyKJkg  : REAL;         // 机房回风比焓 | return air specific enthalpy [kJ/kg]
    rOutdoorTempC        : REAL;         // 户外干球温度 | outdoor dry bulb temperature [℃]
    nUnitsAvail          : INT;          // 可用机组台数 | available unit count [台]
    rDeltaHystKJkg       : REAL := 4.0;  // 焓差滞环半宽 | enthalpy hysteresis half width [kJ/kg]
    rTimeoutS            : REAL := 300.0;// 过渡建立窗（须 ≥120 s，兼作过渡相超时）| transition establish window, also the PARTIAL timeout [s]
END_VAR
VAR_OUTPUT
    nFreeUnits  : INT;                   // 自然冷却投入台数 | units on free cooling [台]
    nMechUnits  : INT;                   // 机械制冷投入台数 | units on mechanical cooling [台]
    xDamperOpen : BOOL;                  // 新风阀开命令（含过渡与混合）| fresh air damper open command, transition and mixed included
    eMode       : E_DL_EconMode;         // 当前模式 | current mode
    xFault      : BOOL;                  // 故障标志 | fault flag
    nFaultCode  : INT;                   // 故障码，锁存至复位沿 | fault code latched until the reset edge
    xActive     : BOOL;                  // 群控已生效回执（未使能时为 FALSE）| group control active acknowledgement
END_VAR
VAR
    tonMech    : TON;                    // MECH 相 最短驻留定时器 | minimum dwell timer of MECH
    tonPartial : TON;                    // PARTIAL 相 建立定时器（阀位渐开）| establish timer of PARTIAL, damper ramping open
    tonFree    : TON;                    // FREE 相 最短驻留定时器 | minimum dwell timer of FREE
    tonMixed   : TON;                    // MIXED 相 最短驻留定时器 | minimum dwell timer of MIXED
    fbEnableFall : F_TRIG;               // xEnable 下降沿（故障复位沿）| falling edge of xEnable, the fault reset edge
    xFinH      : BOOL;                   // 两路比焓有限性 | both enthalpies are finite
    xFinT      : BOOL;                   // 户外温度有限性 | outdoor temperature is finite
    xParamOk   : BOOL;                   // 滞环与超时参数合法 | hysteresis and timeout parameters are legal
    nDwellMs   : UDINT := 120000;        // 最短驻留毫秒数（缺省值防首拍 PT=0）| minimum dwell in milliseconds, default prevents a zero PT
    nPartialMs : UDINT := 300000;        // 过渡建立毫秒数（= rTimeoutS）| transition establish time in milliseconds, equal to rTimeoutS
    xTransCfgOk: BOOL;                   // 过渡配置合法（建立窗 ≥ 最短驻留）| transition configuration legal
    rDiffKJkg  : REAL;                   // 回风比焓 − 户外比焓（正=户外更冷）| return minus outdoor enthalpy, positive when outdoor is cooler [kJ/kg]
    xFreeCond  : BOOL;                   // 全自然冷却条件成立 | free cooling condition satisfied
    xMixedCond : BOOL;                   // 混合冷却条件成立 | mixed cooling condition satisfied
    nHalfUnits : INT;                    // 可用台数的一半 | half of the available units [台]
    nCodeLatch : INT;                    // 故障码锁存副本 | latched copy of the fault code
END_VAR
VAR CONSTANT
    DL_CGE_DWELL_S  : REAL := 120.0;     // 最短驻留时间 | minimum dwell time [s]
    DL_CGE_ENTH_MAX : REAL := 500.0;     // 比焓量程上限 | upper enthalpy range limit [kJ/kg]
    DL_CGE_ENTH_MIN : REAL := -100.0;    // 比焓量程下限 | lower enthalpy range limit [kJ/kg]
    DL_CGE_TEMP_MAX : REAL := 60.0;      // 户外温度量程上限 | upper outdoor temperature limit [℃]
    DL_CGE_TEMP_MIN : REAL := -40.0;     // 户外温度量程下限 | lower outdoor temperature limit [℃]
    DL_CGE_C_NOUNIT : INT := 9601;       // 无可用机组 | no available unit
    DL_CGE_C_ENTH   : INT := 9602;       // 比焓非法 | illegal enthalpy
    DL_CGE_C_TEMP   : INT := 9603;       // 户外温度非法 | illegal outdoor temperature
    DL_CGE_C_TRANS  : INT := 9604;       // 过渡超时 | transition timeout
    DL_CGE_C_UNITS  : INT := 9605;       // 机组数配置越限 | unit count out of range
END_VAR

// 段1｜参数与采样门禁（先判后用，R19：闸断实值通路后再参与比较；换算结果供段2 定时器使用）
xParamOk := (rDeltaHystKJkg = rDeltaHystKJkg) AND ((rDeltaHystKJkg - rDeltaHystKJkg) = 0.0)
            AND (rDeltaHystKJkg >= 0.0)
            AND (rTimeoutS = rTimeoutS) AND ((rTimeoutS - rTimeoutS) = 0.0) AND (rTimeoutS > 0.0);
IF xParamOk THEN
    nPartialMs := REAL_TO_UDINT(rTimeoutS * 1000.0);     // 过渡建立窗 = rTimeoutS（同一参数，避免出现不可达的超时分支）
    nDwellMs := REAL_TO_UDINT(DL_CGE_DWELL_S * 1000.0);
ELSE
    nPartialMs := 300000;                // 参数非法取保守值 | conservative value on an illegal parameter
    nDwellMs := 120000;
END_IF
// 过渡建立窗必须不短于最短驻留，否则自然冷却无法稳定建立，判配置级故障 9604
IF xParamOk THEN
    xTransCfgOk := rTimeoutS >= DL_CGE_DWELL_S;
ELSE
    xTransCfgOk := FALSE;                // 参数本身非法，配置判据不成立 | the parameter itself is illegal
END_IF
xFinH := (rOutdoorEnthalpyKJkg = rOutdoorEnthalpyKJkg) AND ((rOutdoorEnthalpyKJkg - rOutdoorEnthalpyKJkg) = 0.0)
         AND (rReturnEnthalpyKJkg = rReturnEnthalpyKJkg) AND ((rReturnEnthalpyKJkg - rReturnEnthalpyKJkg) = 0.0);
xFinT := (rOutdoorTempC = rOutdoorTempC) AND ((rOutdoorTempC - rOutdoorTempC) = 0.0);

// 段2｜五只定时器 + 一只边沿实例无条件周期刷新（R7，一相一只实例不跨相复用；PT 取自段1 已换算毫秒值）
tonMech(IN := eMode = E_DL_EconMode.MECH, PT := UDINT_TO_TIME(nDwellMs));
tonPartial(IN := eMode = E_DL_EconMode.PARTIAL, PT := UDINT_TO_TIME(nPartialMs));
tonFree(IN := eMode = E_DL_EconMode.FREE, PT := UDINT_TO_TIME(nDwellMs));
tonMixed(IN := eMode = E_DL_EconMode.MIXED, PT := UDINT_TO_TIME(nDwellMs));
fbEnableFall(CLK := xEnable);

// 段3｜输出预置（唯一预置点，CASE 内只置位）
nFreeUnits := 0;
nMechUnits := 0;
xDamperOpen := FALSE;
xFault := FALSE;
nFaultCode := 0;

// 段4｜全局闸：任一入参非法或机组不可用 → 直接锁故障并回机械侧
// R749 码位分判：非有限比焓 → 9602；非有限户外温度 → 9603；参数本身非法 → 9604；三者不再合并为 9602
IF NOT xFinH THEN
    nCodeLatch := DL_CGE_C_ENTH;                 // 比焓非有限 | enthalpy not finite
    xFault := TRUE;
    nFaultCode := DL_CGE_C_ENTH;
    eMode := E_DL_EconMode.FAULT;
ELSIF NOT xFinT THEN
    nCodeLatch := DL_CGE_C_TEMP;                 // 户外温度非有限 | outdoor temperature not finite
    xFault := TRUE;
    nFaultCode := DL_CGE_C_TEMP;
    eMode := E_DL_EconMode.FAULT;
ELSIF NOT xParamOk THEN
    nCodeLatch := DL_CGE_C_TRANS;                // 滞环/超时参数非法（含 NaN 与非正）| illegal hysteresis or timeout parameter
    xFault := TRUE;
    nFaultCode := DL_CGE_C_TRANS;
    eMode := E_DL_EconMode.FAULT;
ELSIF (rOutdoorEnthalpyKJkg > DL_CGE_ENTH_MAX) OR (rOutdoorEnthalpyKJkg < DL_CGE_ENTH_MIN)
      OR (rReturnEnthalpyKJkg > DL_CGE_ENTH_MAX) OR (rReturnEnthalpyKJkg < DL_CGE_ENTH_MIN) THEN
    nCodeLatch := DL_CGE_C_ENTH;
    xFault := TRUE;
    nFaultCode := DL_CGE_C_ENTH;
    eMode := E_DL_EconMode.FAULT;
ELSIF (rOutdoorTempC > DL_CGE_TEMP_MAX) OR (rOutdoorTempC < DL_CGE_TEMP_MIN) THEN
    nCodeLatch := DL_CGE_C_TEMP;
    xFault := TRUE;
    nFaultCode := DL_CGE_C_TEMP;
    eMode := E_DL_EconMode.FAULT;
ELSIF (NOT xTransCfgOk) THEN
    nCodeLatch := DL_CGE_C_TRANS;                // 过渡配置非法：建立窗短于最短驻留 | illegal transition configuration
    xFault := TRUE;
    nFaultCode := DL_CGE_C_TRANS;
    eMode := E_DL_EconMode.FAULT;
ELSIF (nUnitsAvail <= 0) THEN
    nCodeLatch := DL_CGE_C_NOUNIT;
    xFault := TRUE;
    nFaultCode := DL_CGE_C_NOUNIT;
    eMode := E_DL_EconMode.FAULT;
END_IF

// 段5｜判据：回风比焓 − 户外比焓，滞环半宽 rDeltaHystKJkg（判据与出口同源于原始比焓）
IF xFinH THEN
    rDiffKJkg := rReturnEnthalpyKJkg - rOutdoorEnthalpyKJkg;
    xFreeCond := rDiffKJkg > rDeltaHystKJkg;                     // 户外显著更冷 → 全自然 | outdoor clearly cooler, free cooling
    xMixedCond := ABS(rDiffKJkg) <= rDeltaHystKJkg;              // 焓差落在滞环内 → 混合 | gap inside the hysteresis band, mixed
ELSE
    rDiffKJkg := 0.0;                                            // 非有限时不产生判据值 | no criterion when non-finite
    xFreeCond := FALSE;
    xMixedCond := FALSE;
END_IF

// 段6｜主状态机（ENUM + CASE，ELSE 兜底）
IF eMode <> E_DL_EconMode.FAULT THEN
CASE eMode OF
E_DL_EconMode.MECH:
    // 拍 N：全机械，新风阀关闭；驻留满足且全自然条件成立才允许过渡
    IF tonMech.Q THEN
        IF xFreeCond THEN
            eMode := E_DL_EconMode.PARTIAL;          // 本拍行为：进过渡相（阀位渐开）| enter the transition phase
        ELSIF xMixedCond THEN
            eMode := E_DL_EconMode.MIXED;            // 本拍行为：进混合相 | enter the mixed mode
        END_IF
    END_IF

E_DL_EconMode.PARTIAL:
    // 拍 N：过渡相，新风阀渐开、机械减载；条件消失立刻回机械，否则建立窗到即转出
    IF (NOT xFreeCond) AND (NOT xMixedCond) THEN
        eMode := E_DL_EconMode.MECH;                 // 本拍行为：条件消失回机械 | condition lost, back to mechanical
    ELSIF tonPartial.Q THEN
        IF xFreeCond THEN
            eMode := E_DL_EconMode.FREE;             // 本拍行为：建立完成进全自然 | establishment complete, enter free cooling
        ELSE
            eMode := E_DL_EconMode.MIXED;            // 本拍行为：仅满足混合条件进混合 | only the mixed condition holds
        END_IF
    END_IF

E_DL_EconMode.FREE:
    // 拍 N：全自然冷却，驻留满足后才允许退出
    IF tonFree.Q THEN
        IF xMixedCond THEN
            eMode := E_DL_EconMode.MIXED;            // 本拍行为：焓差缩小进混合 | enthalpy gap narrowed, enter mixed
        ELSIF (NOT xFreeCond) AND (NOT xMixedCond) THEN
            eMode := E_DL_EconMode.MECH;             // 本拍行为：条件消失回机械 | back to mechanical
        END_IF
    END_IF

E_DL_EconMode.MIXED:
    // 拍 N：混合冷却，驻留满足后才允许退出
    IF tonMixed.Q THEN
        IF xFreeCond THEN
            eMode := E_DL_EconMode.PARTIAL;          // 本拍行为：焓差放大经过渡进全自然 | gap widened, go through transition
        ELSIF (NOT xFreeCond) AND (NOT xMixedCond) THEN
            eMode := E_DL_EconMode.MECH;             // 本拍行为：条件消失回机械 | back to mechanical
        END_IF
    END_IF

E_DL_EconMode.FAULT:
    // 故障相（本段被外层 IF 排除，保留分支以满足穷举）
    xFault := TRUE;
    nFaultCode := nCodeLatch;

ELSE
    // 非法模式兜底：绝不停在未知模式
    nCodeLatch := DL_CGE_C_UNITS;
    xFault := TRUE;
    nFaultCode := DL_CGE_C_UNITS;
    eMode := E_DL_EconMode.FAULT;
END_CASE
END_IF

// 段7｜每模式独立使能出口与机组分配（故障与兜底一律回机械侧）
// R750 使能门：群控未使能时不得下发任何机组台数与阀位（此前 xEnable 只当复位沿用，名实不符）
IF NOT xEnable THEN
    nFreeUnits := 0;                             // 未使能：自然冷却零台 | disabled, no free cooling unit
    nMechUnits := 0;                             // 未使能：机械侧也零台，交由就地控制 | disabled, no mechanical unit either
    xDamperOpen := FALSE;                        // 未使能：新风阀关 | disabled, damper closed
    xActive := FALSE;                            // 未使能回执 | inactive acknowledgement
ELSE
xActive := TRUE;                                 // 已使能回执 | active acknowledgement
CASE eMode OF
E_DL_EconMode.MECH:
    nFreeUnits := 0;                             // 全机械：无自然冷却台数 | no free cooling units
    nMechUnits := nUnitsAvail;                   // 全机械：可用台数全投 | every available unit on mechanical
    xDamperOpen := FALSE;                        // 新风阀关闭 | damper closed
E_DL_EconMode.PARTIAL:
    nFreeUnits := 1;                             // 过渡：单台先投自然冷却 | one unit on free cooling first
    nMechUnits := nUnitsAvail - nFreeUnits;      // 其余保持机械 | the rest stays mechanical
    xDamperOpen := TRUE;                         // 过渡相独立使能出口：新风阀开 | independent enable of PARTIAL
E_DL_EconMode.FREE:
    nFreeUnits := nUnitsAvail;                   // 全自然：可用台数全投 | every available unit on free cooling
    nMechUnits := 0;
    xDamperOpen := TRUE;                         // 全自然相独立使能出口 | independent enable of FREE
E_DL_EconMode.MIXED:
    nHalfUnits := nUnitsAvail / 2;               // 半数为自然冷却（整数除法，nUnitsAvail 已保证 >0）| half on free cooling
    IF nHalfUnits < 1 THEN
        nHalfUnits := 1;                         // 至少一台，避免混合相退化为全机械 | at least one unit
    END_IF
    nFreeUnits := nHalfUnits;
    nMechUnits := nUnitsAvail - nFreeUnits;
    xDamperOpen := TRUE;                         // 混合相独立使能出口 | independent enable of MIXED
ELSE
    nFreeUnits := 0;                             // 故障与兜底：全机械（安全侧）| fault and fallback, mechanical safe side
    IF nUnitsAvail > 0 THEN
        nMechUnits := nUnitsAvail;               // 机组数有效才下发 | dispatch only a legal unit count
    ELSE
        nMechUnits := 0;                         // 机组数非法不下发负台数（R751）| never dispatch a negative unit count
    END_IF
    xDamperOpen := FALSE;
END_CASE
END_IF

// 段8｜故障相锁存回放与复位沿
IF eMode = E_DL_EconMode.FAULT THEN
    xFault := TRUE;
    nFaultCode := nCodeLatch;                    // 锁存回放，不按当下输入重推断 | republish the latch
    nFreeUnits := 0;                             // 故障相出口强制安全值 | fault outputs forced to the safe side
    IF xEnable AND (nUnitsAvail > 0) THEN
        nMechUnits := nUnitsAvail;               // 已使能且机组数有效：回机械侧安全运行 | enabled with a legal count, run on the mechanical side
    ELSE
        nMechUnits := 0;                         // 未使能或机组数非法：不下发任何台数（R750/R751）| disabled or illegal count, dispatch nothing
    END_IF
    xDamperOpen := FALSE;
    IF fbEnableFall.Q THEN
        nCodeLatch := 0;                         // 清除边：xEnable 下降沿（头注释已声明）| clear edge declared in the header
        eMode := E_DL_EconMode.MECH;
    END_IF
END_IF
END_FUNCTION_BLOCK
